   // ---------- 网络 7 ----------
   // 标题：Z06---> 摄像头防尘盖气缸
   // 注释：临时替换为RSP开关气缸
   // 含义：当 #ST01.Z06.RetEVT 为 TRUE 时置位 #ST01.Z06.IRetPos，否则复位（触点→线圈）
   IF #ST01.Z06.RetEVT THEN
       #ST01.Z06.IRetPos := TRUE;
   ELSE
       #ST01.Z06.IRetPos := FALSE;
   END_IF;
   // 含义：当 #ST01.Z06.ExtEVT 为 TRUE 时置位 #ST01.Z06.IExtPos，否则复位（触点→线圈）
   IF #ST01.Z06.ExtEVT THEN
       #ST01.Z06.IExtPos := TRUE;
   ELSE
       #ST01.Z06.IExtPos := FALSE;
   END_IF;
   // 含义：将 (NOT (#ST01.Z06.ExtEVT) AND #ST01.Z06.IRetPos) AND NOT (#ST01.Z06.IExtPos) 赋给 #ST01.Z06.RetPos
   #ST01.Z06.RetPos := (NOT (#ST01.Z06.ExtEVT) AND #ST01.Z06.IRetPos) AND NOT (#ST01.Z06.IExtPos);
   // 含义：将 (NOT (#ST01.Z06.ExtEVT) AND #ST01.Z06.IRetPos) AND NOT (#ST01.Z06.IExtPos) 赋给 "DB1900_Communication_PC".Send.Z06RetPos
   "DB1900_Communication_PC".Send.Z06RetPos := (NOT (#ST01.Z06.ExtEVT) AND #ST01.Z06.IRetPos) AND NOT (#ST01.Z06.IExtPos);
   // 含义：将 (NOT (#ST01.Z06.RetEVT) AND NOT (#ST01.Z06.IRetPos)) AND #ST01.Z06.IExtPos 赋给 #ST01.Z06.ExtPos
   #ST01.Z06.ExtPos := (NOT (#ST01.Z06.RetEVT) AND NOT (#ST01.Z06.IRetPos)) AND #ST01.Z06.IExtPos;
   // 含义：将 (NOT (#ST01.Z06.RetEVT) AND NOT (#ST01.Z06.IRetPos)) AND #ST01.Z06.IExtPos 赋给 "DB1900_Communication_PC".Send.Z06ExtPos
   "DB1900_Communication_PC".Send.Z06ExtPos := (NOT (#ST01.Z06.RetEVT) AND NOT (#ST01.Z06.IRetPos)) AND #ST01.Z06.IExtPos;
   // 含义：当 #OverAllPmt 为 TRUE 时置位 #ST01.Z06.ExtPmt，否则复位（触点→线圈）
   IF #OverAllPmt THEN
       #ST01.Z06.ExtPmt := TRUE;
   ELSE
       #ST01.Z06.ExtPmt := FALSE;
   END_IF;
   // 含义：当 #OverAllPmt 为 TRUE 时置位 #ST01.Z06.RetPmt，否则复位（触点→线圈）
   IF #OverAllPmt THEN
       #ST01.Z06.RetPmt := TRUE;
   ELSE
       #ST01.Z06.RetPmt := FALSE;
   END_IF;
   // 含义：调用块/实例 "DB1200_FB_std_Switch"，参数：CylinderCmd := #ST01.Z06
   "DB1200_FB_std_Switch"(CylinderCmd := #ST01.Z06);
   // 含义：当 #ST01.Z06.ExtIng 为 TRUE 时置位 "DB1146_PromptFree".ST01.Z06Exting，否则复位（触点→线圈）
   IF #ST01.Z06.ExtIng THEN
       "DB1146_PromptFree".ST01.Z06Exting := TRUE;
   ELSE
       "DB1146_PromptFree".ST01.Z06Exting := FALSE;
   END_IF;
   // 含义：当 #ST01.Z06.RetIng 为 TRUE 时置位 "DB1146_PromptFree".ST01.Z06Reting，否则复位（触点→线圈）
   IF #ST01.Z06.RetIng THEN
       "DB1146_PromptFree".ST01.Z06Reting := TRUE;
   ELSE
       "DB1146_PromptFree".ST01.Z06Reting := FALSE;
   END_IF;
   // 含义：当 #ST01.Z06.ExtErr 为 TRUE 时置位 "DB1148_PromptBeeper".ST01.Z06ExtErr，否则复位（触点→线圈）
   IF #ST01.Z06.ExtErr THEN
       "DB1148_PromptBeeper".ST01.Z06ExtErr := TRUE;
   ELSE
       "DB1148_PromptBeeper".ST01.Z06ExtErr := FALSE;
   END_IF;
   // 含义：当 #ST01.Z06.RetErr 为 TRUE 时置位 "DB1148_PromptBeeper".ST01.Z06RetErr，否则复位（触点→线圈）
   IF #ST01.Z06.RetErr THEN
       "DB1148_PromptBeeper".ST01.Z06RetErr := TRUE;
   ELSE
       "DB1148_PromptBeeper".ST01.Z06RetErr := FALSE;
   END_IF;
   // 含义：条件 "ManMode_M" AND "DB1900_Communication_PC".Recv.Z06ExtTPPB 成立时，将 TRUE 传送到 #ST01.Z06.ExtAuto
   IF "ManMode_M" AND "DB1900_Communication_PC".Recv.Z06ExtTPPB THEN
       #ST01.Z06.ExtAuto := TRUE;
   END_IF;
   // 含义：条件 "ManMode_M" AND "DB1900_Communication_PC".Recv.Z06RetTPPB 成立时，将 TRUE 传送到 #ST01.Z06.RetAuto
   IF "ManMode_M" AND "DB1900_Communication_PC".Recv.Z06RetTPPB THEN
       #ST01.Z06.RetAuto := TRUE;
   END_IF;

   // ---------- 网络 8 ----------
   // 标题：Z07--->快换盘锁紧
   // 含义：将 "IZ07RetPos" AND #Time.ST01Z07RET.Q 赋给 #ST01.Z07.IRetPos
   #ST01.Z07.IRetPos := "IZ07RetPos" AND #Time.ST01Z07RET.Q;
   // 含义：调用定时器实例 #Time.ST01Z07RET.TON
   #Time.ST01Z07RET.TON(IN := "IZ07RetPos",
                        PT := T#1S);
   // 含义：将 "IZ07ExtPos" AND #Time.ST01Z07EXT.Q 赋给 #ST01.Z07.IExtPos
   #ST01.Z07.IExtPos := "IZ07ExtPos" AND #Time.ST01Z07EXT.Q;
   // 含义：调用定时器实例 #Time.ST01Z07EXT.TON
   #Time.ST01Z07EXT.TON(IN := "IZ07ExtPos",
                        PT := T#1S);
   // 含义：将 (NOT (#ST01.Z07.ExtEVT) AND #ST01.Z07.IRetPos) AND NOT (#ST01.Z07.IExtPos) 赋给 #ST01.Z07.RetPos
   #ST01.Z07.RetPos := (NOT (#ST01.Z07.ExtEVT) AND #ST01.Z07.IRetPos) AND NOT (#ST01.Z07.IExtPos);
   // 含义：将 (NOT (#ST01.Z07.ExtEVT) AND #ST01.Z07.IRetPos) AND NOT (#ST01.Z07.IExtPos) 赋给 "DB1900_Communication_PC".Send.Z07RetPos
   "DB1900_Communication_PC".Send.Z07RetPos := (NOT (#ST01.Z07.ExtEVT) AND #ST01.Z07.IRetPos) AND NOT (#ST01.Z07.IExtPos);
   // 含义：将 (NOT (#ST01.Z07.RetEVT) AND NOT (#ST01.Z07.IRetPos)) AND #ST01.Z07.IExtPos 赋给 #ST01.Z07.ExtPos
   #ST01.Z07.ExtPos := (NOT (#ST01.Z07.RetEVT) AND NOT (#ST01.Z07.IRetPos)) AND #ST01.Z07.IExtPos;
   // 含义：将 (NOT (#ST01.Z07.RetEVT) AND NOT (#ST01.Z07.IRetPos)) AND #ST01.Z07.IExtPos 赋给 "DB1900_Communication_PC".Send.Z07ExtPos
   "DB1900_Communication_PC".Send.Z07ExtPos := (NOT (#ST01.Z07.RetEVT) AND NOT (#ST01.Z07.IRetPos)) AND #ST01.Z07.IExtPos;
   // 含义：将 (#OverAllPmt AND "DB720_KuKa_MainCtrl".StatusIn.do_ChgGrp_Pos) OR (#OverAllPmt AND TRUE) 赋给 #ST01.Z07.ExtPmt
   #ST01.Z07.ExtPmt := (#OverAllPmt AND "DB720_KuKa_MainCtrl".StatusIn.do_ChgGrp_Pos) OR (#OverAllPmt AND TRUE);
   // 含义：将 (#OverAllPmt AND "DB720_KuKa_MainCtrl".StatusIn.do_ChgGrp_Pos) OR (#OverAllPmt AND TRUE) 赋给 #ST01.Z07.RetPmt
   #ST01.Z07.RetPmt := (#OverAllPmt AND "DB720_KuKa_MainCtrl".StatusIn.do_ChgGrp_Pos) OR (#OverAllPmt AND TRUE);
   // 含义：调用块/实例 "DB1200_FB_std_Switch"，参数：CylinderCmd := #ST01.Z07
   "DB1200_FB_std_Switch"(CylinderCmd := #ST01.Z07);
   // 含义：当 #ST01.Z07.ExtIng 为 TRUE 时置位 "DB1146_PromptFree".ST01.Z07Exting，否则复位（触点→线圈）
   IF #ST01.Z07.ExtIng THEN
       "DB1146_PromptFree".ST01.Z07Exting := TRUE;
   ELSE
       "DB1146_PromptFree".ST01.Z07Exting := FALSE;
   END_IF;
   // 含义：当 #ST01.Z07.RetIng 为 TRUE 时置位 "DB1146_PromptFree".ST01.Z07Reting，否则复位（触点→线圈）
   IF #ST01.Z07.RetIng THEN
       "DB1146_PromptFree".ST01.Z07Reting := TRUE;
   ELSE
       "DB1146_PromptFree".ST01.Z07Reting := FALSE;
   END_IF;
   // 含义：当 #ST01.Z07.ExtErr 为 TRUE 时置位 "DB1148_PromptBeeper".ST01.Z07ExtErr，否则复位（触点→线圈）
   IF #ST01.Z07.ExtErr THEN
       "DB1148_PromptBeeper".ST01.Z07ExtErr := TRUE;
   ELSE
       "DB1148_PromptBeeper".ST01.Z07ExtErr := FALSE;
   END_IF;
   // 含义：当 #ST01.Z07.RetErr 为 TRUE 时置位 "DB1148_PromptBeeper".ST01.Z07RetErr，否则复位（触点→线圈）
   IF #ST01.Z07.RetErr THEN
       "DB1148_PromptBeeper".ST01.Z07RetErr := TRUE;
   ELSE
       "DB1148_PromptBeeper".ST01.Z07RetErr := FALSE;
   END_IF;
   // 含义：当 #ST01.Z07.ExtEVT 为 TRUE 时置位 "QZ07ExtEvt"，否则复位（触点→线圈）
   IF #ST01.Z07.ExtEVT THEN
       "QZ07ExtEvt" := TRUE;
   ELSE
       "QZ07ExtEvt" := FALSE;
   END_IF;
   // 含义：当 #ST01.Z07.RetEVT 为 TRUE 时置位 "QZ07RetEvt"，否则复位（触点→线圈）
   IF #ST01.Z07.RetEVT THEN
       "QZ07RetEvt" := TRUE;
   ELSE
       "QZ07RetEvt" := FALSE;
   END_IF;
   // 含义：条件 "ManMode_M" AND "DB1900_Communication_PC".Recv.Z07RetTPPB 成立时，将 TRUE 传送到 #ST01.Z07.RetAuto
   IF "ManMode_M" AND "DB1900_Communication_PC".Recv.Z07RetTPPB THEN
       #ST01.Z07.RetAuto := TRUE;
   END_IF;
   // 含义：条件 "ManMode_M" AND "DB1900_Communication_PC".Recv.Z07ExtTPPB 成立时，将 TRUE 传送到 #ST01.Z07.ExtAuto
   IF "ManMode_M" AND "DB1900_Communication_PC".Recv.Z07ExtTPPB THEN
       #ST01.Z07.ExtAuto := TRUE;
   END_IF;

   // ---------- 网络 9 ----------
   // 标题：Z08--->参数写入
   // 含义：将 #ST01.Z08.RetEVT AND #Time.ST01Z08RET.Q 赋给 #ST01.Z08.IRetPos
   #ST01.Z08.IRetPos := #ST01.Z08.RetEVT AND #Time.ST01Z08RET.Q;
   // 含义：调用定时器实例 #Time.ST01Z08RET.TON
   #Time.ST01Z08RET.TON(IN := #ST01.Z08.RetEVT,
                        PT := T#1S);
   // 含义：将 #ST01.Z08.ExtEVT AND #Time.ST01Z08EXT.Q 赋给 #ST01.Z08.IExtPos
   #ST01.Z08.IExtPos := #ST01.Z08.ExtEVT AND #Time.ST01Z08EXT.Q;
   // 含义：调用定时器实例 #Time.ST01Z08EXT.TON
   #Time.ST01Z08EXT.TON(IN := #ST01.Z08.ExtEVT,
                        PT := T#1S);
   // 含义：将 (NOT (#ST01.Z08.ExtEVT) AND #ST01.Z08.IRetPos) AND NOT (#ST01.Z08.IExtPos) 赋给 #ST01.Z08.RetPos
   #ST01.Z08.RetPos := (NOT (#ST01.Z08.ExtEVT) AND #ST01.Z08.IRetPos) AND NOT (#ST01.Z08.IExtPos);
   // 含义：将 (NOT (#ST01.Z08.RetEVT) AND NOT (#ST01.Z08.IRetPos)) AND #ST01.Z08.IExtPos 赋给 #ST01.Z08.ExtPos
   #ST01.Z08.ExtPos := (NOT (#ST01.Z08.RetEVT) AND NOT (#ST01.Z08.IRetPos)) AND #ST01.Z08.IExtPos;
   // 含义：当 #OverAllPmt 为 TRUE 时置位 #ST01.Z08.ExtPmt，否则复位（触点→线圈）
   IF #OverAllPmt THEN
       #ST01.Z08.ExtPmt := TRUE;
   ELSE
       #ST01.Z08.ExtPmt := FALSE;
   END_IF;
   // 含义：当 #OverAllPmt 为 TRUE 时置位 #ST01.Z08.RetPmt，否则复位（触点→线圈）
   IF #OverAllPmt THEN
       #ST01.Z08.RetPmt := TRUE;
   ELSE
       #ST01.Z08.RetPmt := FALSE;
   END_IF;
   // 含义：调用块/实例 "DB1200_FB_std_Switch"，参数：CylinderCmd := #ST01.Z08
   "DB1200_FB_std_Switch"(CylinderCmd := #ST01.Z08);
   // 含义：当 #ST01.Z08.ExtIng 为 TRUE 时置位 "DB1146_PromptFree".ST01.Z08Exting，否则复位（触点→线圈）
   IF #ST01.Z08.ExtIng THEN
       "DB1146_PromptFree".ST01.Z08Exting := TRUE;
   ELSE
       "DB1146_PromptFree".ST01.Z08Exting := FALSE;
   END_IF;
   // 含义：当 #ST01.Z08.RetIng 为 TRUE 时置位 "DB1146_PromptFree".ST01.Z08Reting，否则复位（触点→线圈）
   IF #ST01.Z08.RetIng THEN
       "DB1146_PromptFree".ST01.Z08Reting := TRUE;
   ELSE
       "DB1146_PromptFree".ST01.Z08Reting := FALSE;
   END_IF;
   // 含义：当 #ST01.Z08.ExtErr 为 TRUE 时置位 "DB1148_PromptBeeper".ST01.Z08ExtErr，否则复位（触点→线圈）
   IF #ST01.Z08.ExtErr THEN
       "DB1148_PromptBeeper".ST01.Z08ExtErr := TRUE;
   ELSE
       "DB1148_PromptBeeper".ST01.Z08ExtErr := FALSE;
   END_IF;
   // 含义：当 #ST01.Z08.RetErr 为 TRUE 时置位 "DB1148_PromptBeeper".ST01.Z08RetErr，否则复位（触点→线圈）
   IF #ST01.Z08.RetErr THEN
       "DB1148_PromptBeeper".ST01.Z08RetErr := TRUE;
   ELSE
       "DB1148_PromptBeeper".ST01.Z08RetErr := FALSE;
   END_IF;
   // 含义：当 #ST01.Z08.ExtEVT 为 TRUE 时置位 "DB1900_Communication_PC".Send.ParaWrite，否则复位（触点→线圈）
   IF #ST01.Z08.ExtEVT THEN
       "DB1900_Communication_PC".Send.ParaWrite := TRUE;
   ELSE
       "DB1900_Communication_PC".Send.ParaWrite := FALSE;
   END_IF;
   // 含义：条件 "DB1900_Communication_PC".Recv.ParaWriteDone AND NOT ("ASMMode_M") 成立时，将 TRUE 传送到 #ST01.Z08.RetAuto
   IF "DB1900_Communication_PC".Recv.ParaWriteDone AND NOT ("ASMMode_M") THEN
       #ST01.Z08.RetAuto := TRUE;
   END_IF;
   // 含义：条件 NOT (TRUE) AND NOT ("AllMode_M") 成立时，将 TRUE 传送到 #ST01.Z08.RetAuto
   IF NOT (TRUE) AND NOT ("AllMode_M") THEN
       #ST01.Z08.RetAuto := TRUE;
   END_IF;

   // ---------- 网络 10 ----------
   // 标题：Z09--->三爪卡盘夹爪气缸
   // 含义：条件 (((((NOT (TRUE) AND "AutoMode_M") AND "DB1900_Communication_PC".Para.DrillDirection1) OR ((NOT (TRUE) AND "AutoMode_M") AND "DB1900_Communication_PC".Para.DrillDirection3)) AND NOT ("DB1900_Communication_PC".Para.ProduceMode3)) OR (((((NOT (TRUE) AND "AutoMode_M") AND "DB1900_Communication_PC".Para.DrillDirection1) OR ((NOT (TRUE) AND "AutoMode_M") AND "DB1900_Communication_PC".Para.DrillDirection3)) AND "DB1900_Communication_PC".Para.ProduceMode3) AND "DB1060_AutoStep".HorDrillAutoStep.HorDrillStep.StopDrill_End) OR (((((NOT (TRUE) AND "AutoMode_M") AND "DB1900_Communication_PC".Para.DrillDirection1) OR ((NOT (TRUE) AND "AutoMode_M") AND "DB1900_Communication_PC".Para.DrillDirection3)) AND "DB1900_Communication_PC".Para.ProduceMode3) AND "DB1060_AutoStep".DownDrillAutoStep.DownDrillStep.StopDrill_End)) AND "DB720_KuKa_MainCtrl".Aux.ToolAtPosTimer.Q 成立时，将 TRUE 传送到 #ST01.Z09.ExtEVT
   IF (((((NOT (TRUE) AND "AutoMode_M") AND "DB1900_Communication_PC".Para.DrillDirection1) OR ((NOT (TRUE) AND "AutoMode_M") AND "DB1900_Communication_PC".Para.DrillDirection3)) AND NOT ("DB1900_Communication_PC".Para.ProduceMode3)) OR (((((NOT (TRUE) AND "AutoMode_M") AND "DB1900_Communication_PC".Para.DrillDirection1) OR ((NOT (TRUE) AND "AutoMode_M") AND "DB1900_Communication_PC".Para.DrillDirection3)) AND "DB1900_Communication_PC".Para.ProduceMode3) AND "DB1060_AutoStep".HorDrillAutoStep.HorDrillStep.StopDrill_End) OR (((((NOT (TRUE) AND "AutoMode_M") AND "DB1900_Communication_PC".Para.DrillDirection1) OR ((NOT (TRUE) AND "AutoMode_M") AND "DB1900_Communication_PC".Para.DrillDirection3)) AND "DB1900_Communication_PC".Para.ProduceMode3) AND "DB1060_AutoStep".DownDrillAutoStep.DownDrillStep.StopDrill_End)) AND "DB720_KuKa_MainCtrl".Aux.ToolAtPosTimer.Q THEN
       #ST01.Z09.ExtEVT := TRUE;
   END_IF;
   // 含义：条件 (((((NOT (TRUE) AND "AutoMode_M") AND "DB1900_Communication_PC".Para.DrillDirection1) OR ((NOT (TRUE) AND "AutoMode_M") AND "DB1900_Communication_PC".Para.DrillDirection3)) AND NOT ("DB1900_Communication_PC".Para.ProduceMode3)) OR (((((NOT (TRUE) AND "AutoMode_M") AND "DB1900_Communication_PC".Para.DrillDirection1) OR ((NOT (TRUE) AND "AutoMode_M") AND "DB1900_Communication_PC".Para.DrillDirection3)) AND "DB1900_Communication_PC".Para.ProduceMode3) AND "DB1060_AutoStep".HorDrillAutoStep.HorDrillStep.StopDrill_End) OR (((((NOT (TRUE) AND "AutoMode_M") AND "DB1900_Communication_PC".Para.DrillDirection1) OR ((NOT (TRUE) AND "AutoMode_M") AND "DB1900_Communication_PC".Para.DrillDirection3)) AND "DB1900_Communication_PC".Para.ProduceMode3) AND "DB1060_AutoStep".DownDrillAutoStep.DownDrillStep.StopDrill_End)) AND "DB720_KuKa_MainCtrl".Aux.ToolAtPosTimer.Q 成立时，将 FALSE 传送到 #ST01.Z09.RetEVT
   IF (((((NOT (TRUE) AND "AutoMode_M") AND "DB1900_Communication_PC".Para.DrillDirection1) OR ((NOT (TRUE) AND "AutoMode_M") AND "DB1900_Communication_PC".Para.DrillDirection3)) AND NOT ("DB1900_Communication_PC".Para.ProduceMode3)) OR (((((NOT (TRUE) AND "AutoMode_M") AND "DB1900_Communication_PC".Para.DrillDirection1) OR ((NOT (TRUE) AND "AutoMode_M") AND "DB1900_Communication_PC".Para.DrillDirection3)) AND "DB1900_Communication_PC".Para.ProduceMode3) AND "DB1060_AutoStep".HorDrillAutoStep.HorDrillStep.StopDrill_End) OR (((((NOT (TRUE) AND "AutoMode_M") AND "DB1900_Communication_PC".Para.DrillDirection1) OR ((NOT (TRUE) AND "AutoMode_M") AND "DB1900_Communication_PC".Para.DrillDirection3)) AND "DB1900_Communication_PC".Para.ProduceMode3) AND "DB1060_AutoStep".DownDrillAutoStep.DownDrillStep.StopDrill_End)) AND "DB720_KuKa_MainCtrl".Aux.ToolAtPosTimer.Q THEN
       #ST01.Z09.RetEVT := FALSE;
   END_IF;
   // 含义：调用计数器实例 #Time.ST01Z09EXT.TON（上升沿计数，当前值写入 CV）
   #Time.ST01Z09EXT.TON(IN := (((((((NOT (TRUE) AND "AutoMode_M") AND "DB1900_Communication_PC".Para.DrillDirection1) OR ((NOT (TRUE) AND "AutoMode_M") AND "DB1900_Communication_PC".Para.DrillDirection3)) AND "DB1900_Communication_PC".Para.ProduceMode3) AND "DB720_KuKa_MainCtrl".StatusIn.do_Gouge_Pos) OR (((((NOT (TRUE) AND "AutoMode_M") AND "DB1900_Communication_PC".Para.DrillDirection1) OR ((NOT (TRUE) AND "AutoMode_M") AND "DB1900_Communication_PC".Para.DrillDirection3)) AND "DB1900_Communication_PC".Para.ProduceMode3) AND "DB720_KuKa_MainCtrl".StatusIn.do_DownDril_Pos)) AND ("DB1900_Communication_PC".Recv.Current_2 >= "DB1900_Communication_PC".Para.CurrentMinLimit)),
                        PT := T#30ms);
   // 含义：条件 ((((((NOT (TRUE) AND "AutoMode_M") AND "DB1900_Communication_PC".Para.DrillDirection1) OR ((NOT (TRUE) AND "AutoMode_M") AND "DB1900_Communication_PC".Para.DrillDirection3)) AND "DB1900_Communication_PC".Para.ProduceMode3) AND "DB720_KuKa_MainCtrl".StatusIn.do_Gouge_Pos) OR (((((NOT (TRUE) AND "AutoMode_M") AND "DB1900_Communication_PC".Para.DrillDirection1) OR ((NOT (TRUE) AND "AutoMode_M") AND "DB1900_Communication_PC".Para.DrillDirection3)) AND "DB1900_Communication_PC".Para.ProduceMode3) AND "DB720_KuKa_MainCtrl".StatusIn.do_DownDril_Pos)) AND #Time.ST01Z09EXT.Q 成立时，将 FALSE 传送到 #ST01.Z09.ExtEVT
   IF ((((((NOT (TRUE) AND "AutoMode_M") AND "DB1900_Communication_PC".Para.DrillDirection1) OR ((NOT (TRUE) AND "AutoMode_M") AND "DB1900_Communication_PC".Para.DrillDirection3)) AND "DB1900_Communication_PC".Para.ProduceMode3) AND "DB720_KuKa_MainCtrl".StatusIn.do_Gouge_Pos) OR (((((NOT (TRUE) AND "AutoMode_M") AND "DB1900_Communication_PC".Para.DrillDirection1) OR ((NOT (TRUE) AND "AutoMode_M") AND "DB1900_Communication_PC".Para.DrillDirection3)) AND "DB1900_Communication_PC".Para.ProduceMode3) AND "DB720_KuKa_MainCtrl".StatusIn.do_DownDril_Pos)) AND #Time.ST01Z09EXT.Q THEN
       #ST01.Z09.ExtEVT := FALSE;
   END_IF;
   // 含义：条件 ((((((NOT (TRUE) AND "AutoMode_M") AND "DB1900_Communication_PC".Para.DrillDirection1) OR ((NOT (TRUE) AND "AutoMode_M") AND "DB1900_Communication_PC".Para.DrillDirection3)) AND "DB1900_Communication_PC".Para.ProduceMode3) AND "DB720_KuKa_MainCtrl".StatusIn.do_Gouge_Pos) OR (((((NOT (TRUE) AND "AutoMode_M") AND "DB1900_Communication_PC".Para.DrillDirection1) OR ((NOT (TRUE) AND "AutoMode_M") AND "DB1900_Communication_PC".Para.DrillDirection3)) AND "DB1900_Communication_PC".Para.ProduceMode3) AND "DB720_KuKa_MainCtrl".StatusIn.do_DownDril_Pos)) AND #Time.ST01Z09EXT.Q 成立时，将 TRUE 传送到 #ST01.Z09.RetEVT
   IF ((((((NOT (TRUE) AND "AutoMode_M") AND "DB1900_Communication_PC".Para.DrillDirection1) OR ((NOT (TRUE) AND "AutoMode_M") AND "DB1900_Communication_PC".Para.DrillDirection3)) AND "DB1900_Communication_PC".Para.ProduceMode3) AND "DB720_KuKa_MainCtrl".StatusIn.do_Gouge_Pos) OR (((((NOT (TRUE) AND "AutoMode_M") AND "DB1900_Communication_PC".Para.DrillDirection1) OR ((NOT (TRUE) AND "AutoMode_M") AND "DB1900_Communication_PC".Para.DrillDirection3)) AND "DB1900_Communication_PC".Para.ProduceMode3) AND "DB720_KuKa_MainCtrl".StatusIn.do_DownDril_Pos)) AND #Time.ST01Z09EXT.Q THEN
       #ST01.Z09.RetEVT := TRUE;
   END_IF;
   // 含义：条件 ((((NOT (TRUE) AND "AutoMode_M") AND "DB1900_Communication_PC".Para.DrillDirection1) OR ((NOT (TRUE) AND "AutoMode_M") AND "DB1900_Communication_PC".Para.DrillDirection3)) AND "DB1900_Communication_PC".Para.ProduceMode3) AND #ST01.Z09.ExtEVT 成立时，将 TRUE 传送到 "QZ14ExtEvt"
   IF ((((NOT (TRUE) AND "AutoMode_M") AND "DB1900_Communication_PC".Para.DrillDirection1) OR ((NOT (TRUE) AND "AutoMode_M") AND "DB1900_Communication_PC".Para.DrillDirection3)) AND "DB1900_Communication_PC".Para.ProduceMode3) AND #ST01.Z09.ExtEVT THEN
       "QZ14ExtEvt" := TRUE;
   END_IF;
   // 含义：条件 ((((NOT (TRUE) AND "AutoMode_M") AND "DB1900_Communication_PC".Para.DrillDirection1) OR ((NOT (TRUE) AND "AutoMode_M") AND "DB1900_Communication_PC".Para.DrillDirection3)) AND "DB1900_Communication_PC".Para.ProduceMode3) AND #ST01.Z09.ExtEVT 成立时，将 FALSE 传送到 "QZ14RetEvt"
   IF ((((NOT (TRUE) AND "AutoMode_M") AND "DB1900_Communication_PC".Para.DrillDirection1) OR ((NOT (TRUE) AND "AutoMode_M") AND "DB1900_Communication_PC".Para.DrillDirection3)) AND "DB1900_Communication_PC".Para.ProduceMode3) AND #ST01.Z09.ExtEVT THEN
       "QZ14RetEvt" := FALSE;
   END_IF;
   // 含义：条件 ((((NOT (TRUE) AND "AutoMode_M") AND "DB1900_Communication_PC".Para.DrillDirection1) OR ((NOT (TRUE) AND "AutoMode_M") AND "DB1900_Communication_PC".Para.DrillDirection3)) AND "DB1900_Communication_PC".Para.ProduceMode3) AND #ST01.Z09.RetEVT 成立时，将 FALSE 传送到 "QZ14ExtEvt"
   IF ((((NOT (TRUE) AND "AutoMode_M") AND "DB1900_Communication_PC".Para.DrillDirection1) OR ((NOT (TRUE) AND "AutoMode_M") AND "DB1900_Communication_PC".Para.DrillDirection3)) AND "DB1900_Communication_PC".Para.ProduceMode3) AND #ST01.Z09.RetEVT THEN
       "QZ14ExtEvt" := FALSE;
   END_IF;
   // 含义：条件 ((((NOT (TRUE) AND "AutoMode_M") AND "DB1900_Communication_PC".Para.DrillDirection1) OR ((NOT (TRUE) AND "AutoMode_M") AND "DB1900_Communication_PC".Para.DrillDirection3)) AND "DB1900_Communication_PC".Para.ProduceMode3) AND #ST01.Z09.RetEVT 成立时，将 TRUE 传送到 "QZ14RetEvt"
   IF ((((NOT (TRUE) AND "AutoMode_M") AND "DB1900_Communication_PC".Para.DrillDirection1) OR ((NOT (TRUE) AND "AutoMode_M") AND "DB1900_Communication_PC".Para.DrillDirection3)) AND "DB1900_Communication_PC".Para.ProduceMode3) AND #ST01.Z09.RetEVT THEN
       "QZ14RetEvt" := TRUE;
   END_IF;
   // 含义：条件 (NOT (TRUE) AND "ManMode_M") OR ((NOT (TRUE) AND "AutoMode_M") AND NOT ("DB1900_Communication_PC".Send.DrillRunning)) 成立时，将 FALSE 传送到 #ST01.Z09.ExtEVT
   IF (NOT (TRUE) AND "ManMode_M") OR ((NOT (TRUE) AND "AutoMode_M") AND NOT ("DB1900_Communication_PC".Send.DrillRunning)) THEN
       #ST01.Z09.ExtEVT := FALSE;
   END_IF;
   // 含义：条件 (NOT (TRUE) AND "ManMode_M") OR ((NOT (TRUE) AND "AutoMode_M") AND NOT ("DB1900_Communication_PC".Send.DrillRunning)) 成立时，将 FALSE 传送到 #ST01.Z09.RetEVT
   IF (NOT (TRUE) AND "ManMode_M") OR ((NOT (TRUE) AND "AutoMode_M") AND NOT ("DB1900_Communication_PC".Send.DrillRunning)) THEN
       #ST01.Z09.RetEVT := FALSE;
   END_IF;

   // ---------- 网络 11 ----------
   // （空白网络）
END_FUNCTION_BLOCK

FUNCTION_BLOCK "FB1910_DrillData"   // FB1910, SCL
{ S7_Optimized_Access := 'TRUE' }
// ============================================================
//  Block: FB1910_DrillData
//  ============================================================
//  编号：FB1910
//  原始语言：LAD（规则翻译为 SCL）
//  含义：Hammer
   VAR
      HorDrill : "UDT_DrillData";   // 水平水泥数据
      DownDrill : "UDT_DrillData";   // 垂直向下水泥数据
      AUX : Struct   // 静态变量
         LayerNo : Int := 1;   // 层数记忆
         HDirection : Int := 1;   // 水平方向1正2负
         DDirection : Int := 1;   // 向下方向1正2负
         GougeDrillWidth : Real;   // 凿击宽度要加10
      END_STRUCT;
      EdgeDetc : Struct   // 静态变量
         Pulse : Array[0..15] of Bool;   // 静态变量
      END_STRUCT;
      CurrentDrillWidth : Real;   // 静态变量
      CurrentDrillLength : Real;   // 静态变量
      CurrentDrillDepth : Real;   // 静态变量
      LastDrillWidth : Real;   // 静态变量
      LastDrillDepth : Real;   // 静态变量
      AlreadyDrillWidth : Real;   // 静态变量
      AlreadyDrillLength : Real;   // 静态变量
      MaxWidth : Real;   // 静态变量
      gi_OffsetX : Real;   // 静态变量
      gi_OffSetY : Real;   // 静态变量
      gi_OffSetZ : Real;   // 静态变量
      SlabWidth : Real := 0.0;   // 静态变量
      SlabLength : Real := 0.0;   // 静态变量
      PosNo : Int;   // 静态变量
      OppositeStartPos : Real;   // 静态变量
   END_VAR
   VAR_TEMP
      HorPosMod : Int;   // 临时变量
      DownPosMod : Int;   // 临时变量
   END_VAR
BEGIN

   // ---------- 网络 1 ----------
   // 标题：水泥长宽输入
   // 含义：条件 ((("DB1900_Communication_PC".Para.HorConcreteZ > 100.0) AND ("DB720_KuKa_MainCtrl".CmdOut.gi_ToolTypeNo = 2))) OR ((("DB1900_Communication_PC".Para.HorConcreteZ > 100.0) AND ("DB720_KuKa_MainCtrl".CmdOut.gi_ToolTypeNo = 18))) 成立时，将 "DB1900_Communication_PC".Para.HorConcreteZ 传送到 #HorDrill.SlabWidth
   IF ((("DB1900_Communication_PC".Para.HorConcreteZ > 100.0) AND ("DB720_KuKa_MainCtrl".CmdOut.gi_ToolTypeNo = 2))) OR ((("DB1900_Communication_PC".Para.HorConcreteZ > 100.0) AND ("DB720_KuKa_MainCtrl".CmdOut.gi_ToolTypeNo = 18))) THEN
       #HorDrill.SlabWidth := "DB1900_Communication_PC".Para.HorConcreteZ;
   END_IF;
   // 含义：条件 (((("DB1900_Communication_PC".Para.HorConcreteZ > 100.0) AND ("DB720_KuKa_MainCtrl".CmdOut.gi_ToolTypeNo = 13))) AND ("DB1900_Communication_PC".Para.Classification = 1)) 成立时，将 500.0 传送到 #HorDrill.SlabWidth
   IF (((("DB1900_Communication_PC".Para.HorConcreteZ > 100.0) AND ("DB720_KuKa_MainCtrl".CmdOut.gi_ToolTypeNo = 13))) AND ("DB1900_Communication_PC".Para.Classification = 1)) THEN
       #HorDrill.SlabWidth := 500.0;
   END_IF;
   // 含义：条件 ((((("DB1900_Communication_PC".Para.HorConcreteZ > 100.0) AND ("DB720_KuKa_MainCtrl".CmdOut.gi_ToolTypeNo = 13))) AND ("DB1900_Communication_PC".Para.Classification = 2))) OR ((((("DB1900_Communication_PC".Para.HorConcreteZ > 100.0) AND ("DB720_KuKa_MainCtrl".CmdOut.gi_ToolTypeNo = 13))) AND ("DB1900_Communication_PC".Para.Classification = 3))) 成立时，将 850.0 传送到 #HorDrill.SlabWidth
   IF ((((("DB1900_Communication_PC".Para.HorConcreteZ > 100.0) AND ("DB720_KuKa_MainCtrl".CmdOut.gi_ToolTypeNo = 13))) AND ("DB1900_Communication_PC".Para.Classification = 2))) OR ((((("DB1900_Communication_PC".Para.HorConcreteZ > 100.0) AND ("DB720_KuKa_MainCtrl".CmdOut.gi_ToolTypeNo = 13))) AND ("DB1900_Communication_PC".Para.Classification = 3))) THEN
       #HorDrill.SlabWidth := 850.0;
   END_IF;
   // 含义：条件 ((("DB1900_Communication_PC".Para.HorConcreteY > 200.0) AND ("DB720_KuKa_MainCtrl".CmdOut.gi_ToolTypeNo = 2))) OR ((("DB1900_Communication_PC".Para.HorConcreteY > 200.0) AND ("DB720_KuKa_MainCtrl".CmdOut.gi_ToolTypeNo = 18))) 成立时，将 "DB1900_Communication_PC".Para.HorConcreteY 传送到 #HorDrill.SlabLength
   IF ((("DB1900_Communication_PC".Para.HorConcreteY > 200.0) AND ("DB720_KuKa_MainCtrl".CmdOut.gi_ToolTypeNo = 2))) OR ((("DB1900_Communication_PC".Para.HorConcreteY > 200.0) AND ("DB720_KuKa_MainCtrl".CmdOut.gi_ToolTypeNo = 18))) THEN
       #HorDrill.SlabLength := "DB1900_Communication_PC".Para.HorConcreteY;
   END_IF;
   // 含义：条件 (((("DB1900_Communication_PC".Para.HorConcreteY > 200.0) AND ("DB720_KuKa_MainCtrl".CmdOut.gi_ToolTypeNo = 13))) AND ("DB1900_Communication_PC".Para.DrillWidth <> 105.0)) 成立时，将 960.0 传送到 #HorDrill.SlabLength
   IF (((("DB1900_Communication_PC".Para.HorConcreteY > 200.0) AND ("DB720_KuKa_MainCtrl".CmdOut.gi_ToolTypeNo = 13))) AND ("DB1900_Communication_PC".Para.DrillWidth <> 105.0)) THEN
       #HorDrill.SlabLength := 960.0;
   END_IF;
   // 含义：条件 (((("DB1900_Communication_PC".Para.HorConcreteY > 200.0) AND ("DB720_KuKa_MainCtrl".CmdOut.gi_ToolTypeNo = 13))) AND ("DB1900_Communication_PC".Para.DrillWidth = 105.0)) 成立时，将 1100.0 传送到 #HorDrill.SlabLength
   IF (((("DB1900_Communication_PC".Para.HorConcreteY > 200.0) AND ("DB720_KuKa_MainCtrl".CmdOut.gi_ToolTypeNo = 13))) AND ("DB1900_Communication_PC".Para.DrillWidth = 105.0)) THEN
       #HorDrill.SlabLength := 1100.0;
   END_IF;
   // 含义：条件 ("DB1900_Communication_PC".Para.DownConcreteX > 50.0) 成立时，将 "DB1900_Communication_PC".Para.DownConcreteX 传送到 #DownDrill.SlabWidth
   IF ("DB1900_Communication_PC".Para.DownConcreteX > 50.0) THEN
       #DownDrill.SlabWidth := "DB1900_Communication_PC".Para.DownConcreteX;
   END_IF;
   // 含义：条件 (("DB1900_Communication_PC".Para.DownConcreteY > 100.0) AND ("DB720_KuKa_MainCtrl".CmdOut.gi_ToolTypeNo = 2)) 成立时，将 "DB1900_Communication_PC".Para.DownConcreteY 传送到 #DownDrill.SlabLength
   IF (("DB1900_Communication_PC".Para.DownConcreteY > 100.0) AND ("DB720_KuKa_MainCtrl".CmdOut.gi_ToolTypeNo = 2)) THEN
       #DownDrill.SlabLength := "DB1900_Communication_PC".Para.DownConcreteY;
   END_IF;
   // 含义：条件 (("DB1900_Communication_PC".Para.DownConcreteY > 100.0) AND ("DB720_KuKa_MainCtrl".CmdOut.gi_ToolTypeNo = 13)) 成立时，将 1110.0 传送到 #DownDrill.SlabLength
   IF (("DB1900_Communication_PC".Para.DownConcreteY > 100.0) AND ("DB720_KuKa_MainCtrl".CmdOut.gi_ToolTypeNo = 13)) THEN
       #DownDrill.SlabLength := 1110.0;
   END_IF;
   // 含义：条件 ("DB1900_Communication_PC".Recv.Layer < 1) 成立时，将 1 传送到 "DB1900_Communication_PC".Recv.Layer
   IF ("DB1900_Communication_PC".Recv.Layer < 1) THEN
       "DB1900_Communication_PC".Recv.Layer := 1;
   END_IF;
   // 含义：条件 "DB1900_Communication_PC".Recv.PowerOff OR ("ManMode_M" AND "ErrRst_M") 成立时，将 FALSE 传送到 "DB1900_Communication_PC".Send.PowerOff
   IF "DB1900_Communication_PC".Recv.PowerOff OR ("ManMode_M" AND "ErrRst_M") THEN
       "DB1900_Communication_PC".Send.PowerOff := FALSE;
   END_IF;

   // ---------- 网络 2 ----------
   // 标题：锤钻打孔长宽输入
   // 注释：Hammer
   // 含义：条件 ((("DB720_KuKa_MainCtrl".CmdOut.gi_ToolTypeNo = 2) OR ("DB720_KuKa_MainCtrl".CmdOut.gi_ToolTypeNo = 18)) AND "DB1900_Communication_PC".Para.DrillDirection1) AND NOT ("DB1900_Communication_PC".Para.ProduceMode3) 成立时，将 "DB1900_Communication_PC".Para.DrillWidth 传送到 #HorDrill.CurrentDrillWidth
   IF ((("DB720_KuKa_MainCtrl".CmdOut.gi_ToolTypeNo = 2) OR ("DB720_KuKa_MainCtrl".CmdOut.gi_ToolTypeNo = 18)) AND "DB1900_Communication_PC".Para.DrillDirection1) AND NOT ("DB1900_Communication_PC".Para.ProduceMode3) THEN
       #HorDrill.CurrentDrillWidth := "DB1900_Communication_PC".Para.DrillWidth;
   END_IF;
   // 含义：条件 ((("DB720_KuKa_MainCtrl".CmdOut.gi_ToolTypeNo = 2) OR ("DB720_KuKa_MainCtrl".CmdOut.gi_ToolTypeNo = 18)) AND "DB1900_Communication_PC".Para.DrillDirection1) AND "DB1900_Communication_PC".Para.ProduceMode3 成立时，将 ("DB1900_Communication_PC".Para.DrillWidth + 10.0) 传送到 #HorDrill.CurrentDrillWidth
   IF ((("DB720_KuKa_MainCtrl".CmdOut.gi_ToolTypeNo = 2) OR ("DB720_KuKa_MainCtrl".CmdOut.gi_ToolTypeNo = 18)) AND "DB1900_Communication_PC".Para.DrillDirection1) AND "DB1900_Communication_PC".Para.ProduceMode3 THEN
       #HorDrill.CurrentDrillWidth := ("DB1900_Communication_PC".Para.DrillWidth + 10.0);
   END_IF;
   // 含义：条件 (("DB720_KuKa_MainCtrl".CmdOut.gi_ToolTypeNo = 2) OR ("DB720_KuKa_MainCtrl".CmdOut.gi_ToolTypeNo = 18)) AND "DB1900_Communication_PC".Para.DrillDirection1 成立时，将 "DB1900_Communication_PC".Para.DrillWidth 传送到 #HorDrill.CurrentDrillLength
   IF (("DB720_KuKa_MainCtrl".CmdOut.gi_ToolTypeNo = 2) OR ("DB720_KuKa_MainCtrl".CmdOut.gi_ToolTypeNo = 18)) AND "DB1900_Communication_PC".Para.DrillDirection1 THEN
       #HorDrill.CurrentDrillLength := "DB1900_Communication_PC".Para.DrillWidth;
   END_IF;
   // 含义：条件 (("DB720_KuKa_MainCtrl".CmdOut.gi_ToolTypeNo = 2) OR ("DB720_KuKa_MainCtrl".CmdOut.gi_ToolTypeNo = 18)) AND "DB1900_Communication_PC".Para.DrillDirection3 成立时，将 "DB1900_Communication_PC".Para.DrillWidth 传送到 #DownDrill.CurrentDrillWidth
   IF (("DB720_KuKa_MainCtrl".CmdOut.gi_ToolTypeNo = 2) OR ("DB720_KuKa_MainCtrl".CmdOut.gi_ToolTypeNo = 18)) AND "DB1900_Communication_PC".Para.DrillDirection3 THEN
       #DownDrill.CurrentDrillWidth := "DB1900_Communication_PC".Para.DrillWidth;
   END_IF;

   // ---------- 网络 3 ----------
   // 标题：打孔水钻长宽输入
   // 注释：Core Diamond Drill
   // 32mm: Hor; Height:  45mm; Length: 50mm 100mm   150mm 250mm
   // 52mm:Down; Height: 65mm; Length: 66.66mm 132.33mmmm   233.67mm
   // 82mm Hor; Height:85mm; Length:100mm 300mm
   // 102mm Hor; Height:80mm; Length:400mm
   // 132mm Hor; Height:120mm; Length:400mm
   // 含义：条件 ((((("DB720_KuKa_MainCtrl".CmdOut.gi_ToolTypeNo = 13) AND "DB1900_Communication_PC".Para.DrillDirection1) AND ("DB1900_Communication_PC".Para.DrillWidth = 45.0))) AND ("DB1900_Communication_PC".Para.Classification = 1)) 成立时，将 (#HorDrill.PosNo MOD 4) 传送到 #HorPosMod
   IF ((((("DB720_KuKa_MainCtrl".CmdOut.gi_ToolTypeNo = 13) AND "DB1900_Communication_PC".Para.DrillDirection1) AND ("DB1900_Communication_PC".Para.DrillWidth = 45.0))) AND ("DB1900_Communication_PC".Para.Classification = 1)) THEN
       #HorPosMod := (#HorDrill.PosNo MOD 4);
   END_IF;
   // 含义：条件 ((#HorDrill.PosNo >= 1) AND (#HorPosMod = 3)) 成立时，将 250.0 传送到 #HorDrill.CurrentDrillLength
   IF ((#HorDrill.PosNo >= 1) AND (#HorPosMod = 3)) THEN
       #HorDrill.CurrentDrillLength := 250.0;
   END_IF;
   // 含义：条件 ((#HorDrill.PosNo >= 1) AND (#HorPosMod <> 3)) 成立时，将 50.0 传送到 #HorDrill.CurrentDrillLength
   IF ((#HorDrill.PosNo >= 1) AND (#HorPosMod <> 3)) THEN
       #HorDrill.CurrentDrillLength := 50.0;
   END_IF;
   // 含义：条件 ((#HorDrill.PosNo = 0) AND (#HorPosMod = 0)) 成立时，将 50.0 传送到 #HorDrill.CurrentDrillLength
   IF ((#HorDrill.PosNo = 0) AND (#HorPosMod = 0)) THEN
       #HorDrill.CurrentDrillLength := 50.0;
   END_IF;
   // 含义：条件 ((((("DB720_KuKa_MainCtrl".CmdOut.gi_ToolTypeNo = 13) AND "DB1900_Communication_PC".Para.DrillDirection1) AND ("DB1900_Communication_PC".Para.DrillWidth = 65.0))) AND ("DB1900_Communication_PC".Para.Classification = 1)) 成立时，将 (#HorDrill.PosNo MOD 3) 传送到 #HorPosMod
   IF ((((("DB720_KuKa_MainCtrl".CmdOut.gi_ToolTypeNo = 13) AND "DB1900_Communication_PC".Para.DrillDirection1) AND ("DB1900_Communication_PC".Para.DrillWidth = 65.0))) AND ("DB1900_Communication_PC".Para.Classification = 1)) THEN
       #HorPosMod := (#HorDrill.PosNo MOD 3);
   END_IF;
   // 含义：条件 ((#HorDrill.PosNo >= 1) AND (#HorPosMod = 2)) 成立时，将 266.68 传送到 #HorDrill.CurrentDrillLength
   IF ((#HorDrill.PosNo >= 1) AND (#HorPosMod = 2)) THEN
       #HorDrill.CurrentDrillLength := 266.68;
   END_IF;
   // 含义：条件 ((#HorDrill.PosNo >= 1) AND (#HorPosMod <> 2)) 成立时，将 66.66 传送到 #HorDrill.CurrentDrillLength
   IF ((#HorDrill.PosNo >= 1) AND (#HorPosMod <> 2)) THEN
       #HorDrill.CurrentDrillLength := 66.66;
   END_IF;
   // 含义：条件 ((#HorDrill.PosNo = 0) AND (#HorPosMod = 0)) 成立时，将 66.66 传送到 #HorDrill.CurrentDrillLength
   IF ((#HorDrill.PosNo = 0) AND (#HorPosMod = 0)) THEN
       #HorDrill.CurrentDrillLength := 66.66;
   END_IF;
   // 含义：条件 (((((("DB720_KuKa_MainCtrl".CmdOut.gi_ToolTypeNo = 13) AND "DB1900_Communication_PC".Para.DrillDirection1) AND ("DB1900_Communication_PC".Para.DrillWidth = 85.0))) AND ("DB1900_Communication_PC".Para.Classification = 2))) OR (((((("DB720_KuKa_MainCtrl".CmdOut.gi_ToolTypeNo = 13) AND "DB1900_Communication_PC".Para.DrillDirection1) AND ("DB1900_Communication_PC".Para.DrillWidth = 85.0))) AND ("DB1900_Communication_PC".Para.Classification = 3))) 成立时，将 (#HorDrill.PosNo MOD 2) 传送到 #HorPosMod
   IF (((((("DB720_KuKa_MainCtrl".CmdOut.gi_ToolTypeNo = 13) AND "DB1900_Communication_PC".Para.DrillDirection1) AND ("DB1900_Communication_PC".Para.DrillWidth = 85.0))) AND ("DB1900_Communication_PC".Para.Classification = 2))) OR (((((("DB720_KuKa_MainCtrl".CmdOut.gi_ToolTypeNo = 13) AND "DB1900_Communication_PC".Para.DrillDirection1) AND ("DB1900_Communication_PC".Para.DrillWidth = 85.0))) AND ("DB1900_Communication_PC".Para.Classification = 3))) THEN
       #HorPosMod := (#HorDrill.PosNo MOD 2);
   END_IF;
   // 含义：条件 ((#HorDrill.PosNo >= 1) AND (#HorPosMod = 1)) 成立时，将 300.0 传送到 #HorDrill.CurrentDrillLength
   IF ((#HorDrill.PosNo >= 1) AND (#HorPosMod = 1)) THEN
       #HorDrill.CurrentDrillLength := 300.0;
   END_IF;
   // 含义：条件 ((#HorDrill.PosNo >= 1) AND (#HorPosMod <> 1)) 成立时，将 100.0 传送到 #HorDrill.CurrentDrillLength
   IF ((#HorDrill.PosNo >= 1) AND (#HorPosMod <> 1)) THEN
       #HorDrill.CurrentDrillLength := 100.0;
   END_IF;
   // 含义：条件 ((#HorDrill.PosNo = 0) AND (#HorPosMod = 0)) 成立时，将 100.0 传送到 #HorDrill.CurrentDrillLength
   IF ((#HorDrill.PosNo = 0) AND (#HorPosMod = 0)) THEN
       #HorDrill.CurrentDrillLength := 100.0;
   END_IF;
   // 含义：条件 ((((("DB720_KuKa_MainCtrl".CmdOut.gi_ToolTypeNo = 13) AND "DB1900_Communication_PC".Para.DrillDirection1) AND ("DB1900_Communication_PC".Para.DrillWidth = 105.0))) AND ("DB1900_Communication_PC".Para.Classification = 1)) 成立时，将 125.0 传送到 #HorDrill.CurrentDrillLength
   IF ((((("DB720_KuKa_MainCtrl".CmdOut.gi_ToolTypeNo = 13) AND "DB1900_Communication_PC".Para.DrillDirection1) AND ("DB1900_Communication_PC".Para.DrillWidth = 105.0))) AND ("DB1900_Communication_PC".Para.Classification = 1)) THEN
       #HorDrill.CurrentDrillLength := 125.0;
   END_IF;
   // 含义：条件 (((((("DB720_KuKa_MainCtrl".CmdOut.gi_ToolTypeNo = 13) AND "DB1900_Communication_PC".Para.DrillDirection1) AND ("DB1900_Communication_PC".Para.DrillWidth = 80.0))) OR (((("DB720_KuKa_MainCtrl".CmdOut.gi_ToolTypeNo = 13) AND "DB1900_Communication_PC".Para.DrillDirection1) AND ("DB1900_Communication_PC".Para.DrillWidth = 120.0)))) AND ("DB1900_Communication_PC".Para.Classification = 2)) 成立时，将 400.0 传送到 #HorDrill.CurrentDrillLength
   IF (((((("DB720_KuKa_MainCtrl".CmdOut.gi_ToolTypeNo = 13) AND "DB1900_Communication_PC".Para.DrillDirection1) AND ("DB1900_Communication_PC".Para.DrillWidth = 80.0))) OR (((("DB720_KuKa_MainCtrl".CmdOut.gi_ToolTypeNo = 13) AND "DB1900_Communication_PC".Para.DrillDirection1) AND ("DB1900_Communication_PC".Para.DrillWidth = 120.0)))) AND ("DB1900_Communication_PC".Para.Classification = 2)) THEN
       #HorDrill.CurrentDrillLength := 400.0;
   END_IF;
   // 含义：条件 ("DB720_KuKa_MainCtrl".CmdOut.gi_ToolTypeNo = 13) AND "DB1900_Communication_PC".Para.DrillDirection1 成立时，将 "DB1900_Communication_PC".Para.DrillWidth 传送到 #HorDrill.CurrentDrillWidth
   IF ("DB720_KuKa_MainCtrl".CmdOut.gi_ToolTypeNo = 13) AND "DB1900_Communication_PC".Para.DrillDirection1 THEN
       #HorDrill.CurrentDrillWidth := "DB1900_Communication_PC".Para.DrillWidth;
   END_IF;
   // 含义：条件 ((("DB720_KuKa_MainCtrl".CmdOut.gi_ToolTypeNo = 13) AND "DB1900_Communication_PC".Para.DrillDirection3) AND ("DB1900_Communication_PC".Para.DrillWidth = 65.0)) 成立时，将 (#DownDrill.PosNo MOD 3) 传送到 #DownPosMod
   IF ((("DB720_KuKa_MainCtrl".CmdOut.gi_ToolTypeNo = 13) AND "DB1900_Communication_PC".Para.DrillDirection3) AND ("DB1900_Communication_PC".Para.DrillWidth = 65.0)) THEN
       #DownPosMod := (#DownDrill.PosNo MOD 3);
   END_IF;
   // 含义：条件 ((#DownDrill.PosNo >= 1) AND (#DownPosMod = 2)) 成立时，将 266.68 传送到 #DownDrill.CurrentDrillLength
   IF ((#DownDrill.PosNo >= 1) AND (#DownPosMod = 2)) THEN
       #DownDrill.CurrentDrillLength := 266.68;
   END_IF;
   // 含义：条件 ((#DownDrill.PosNo >= 1) AND (#DownPosMod <> 2)) 成立时，将 66.6 传送到 #DownDrill.CurrentDrillLength
   IF ((#DownDrill.PosNo >= 1) AND (#DownPosMod <> 2)) THEN
       #DownDrill.CurrentDrillLength := 66.6;
   END_IF;
   // 含义：条件 ((#DownDrill.PosNo = 0) AND (#DownPosMod = 0)) 成立时，将 66.6 传送到 #HorDrill.CurrentDrillLength
   IF ((#DownDrill.PosNo = 0) AND (#DownPosMod = 0)) THEN
       #HorDrill.CurrentDrillLength := 66.6;
   END_IF;
   // 含义：条件 ("DB720_KuKa_MainCtrl".CmdOut.gi_ToolTypeNo = 13) AND "DB1900_Communication_PC".Para.DrillDirection3 成立时，将 "DB1900_Communication_PC".Para.DrillWidth 传送到 #DownDrill.CurrentDrillWidth
   IF ("DB720_KuKa_MainCtrl".CmdOut.gi_ToolTypeNo = 13) AND "DB1900_Communication_PC".Para.DrillDirection3 THEN
       #DownDrill.CurrentDrillWidth := "DB1900_Communication_PC".Para.DrillWidth;
   END_IF;

   // ---------- 网络 4 ----------
   // 标题：手动输入水平水泥数据处理
   // 含义：本网络为 StructuredText（SCL）原文重建，非 LAD 折叠
   IF "DB1900_Communication_PC".Recv.HorizontalConfirm AND "IMan" THEN
       #AUX.HDirection := 1;
       #HorDrill.OppositeStartPos := 0;
       #AUX.LayerNo := "DB1900_Communication_PC".Recv.Layer;
       #HorDrill.LastDrillWidth := #HorDrill.CurrentDrillWidth;
       #HorDrill.gi_OffSetZ := ABS("DB1900_Communication_PC".Recv.Horizontal_OffSetZ);
       #HorDrill.gi_OffSetY := ABS("DB1900_Communication_PC".Recv.Horizontal_OffSetY);
       #HorDrill.AlreadyDrillWidth := ABS("DB1900_Communication_PC".Recv.Horizontal_OffSetZ);
       #HorDrill.AlreadyDrillLength := ABS("DB1900_Communication_PC".Recv.Horizontal_OffSetY);
       IF "DB1900_Communication_PC".Recv.Horizontal_OffSetY = 0 THEN
           #HorDrill.PosNo := 0;
       END_IF;
   END_IF;
   IF "DB1900_Communication_PC".Recv.ChangeHorizontalSlabDone AND "IMan" THEN
       #AUX.LayerNo := 1;
       #AUX.HDirection := 1;
       #HorDrill.PosNo := 0;
       #HorDrill.gi_OffSetZ := 0;
       #HorDrill.gi_OffSetY := 0;
       #HorDrill.OppositeStartPos := 0;
       #HorDrill.AlreadyDrillWidth := 0;
       #HorDrill.AlreadyDrillLength := 0;
       #HorDrill.LastDrillWidth := #HorDrill.CurrentDrillWidth;
       "DB1147_PromptStartNotPmt".Public.ChangeHorDrillSlab := FALSE;
   END_IF;

   // ---------- 网络 5 ----------
   // 标题：水平水泥数据 Y平长 Z纵宽
   // 含义：本网络为 StructuredText（SCL）原文重建，非 LAD 折叠
   IF "DB1900_Communication_PC".Para.DrillDirection1 = TRUE AND (NOT "DB1900_Communication_PC".Para.ProduceMode3) AND "AutoMode_M" THEN
       IF "DB2500 Visual Chiseling".VChiselCamRound = -1 THEN
           #HorDrill.SlabWidth := #HorDrill.SlabWidth;
       ELSIF ("DB2500 Visual Chiseling".VChiselCamRound >= 0 AND "DB2500 Visual Chiseling".VChiselCamRound <= 44) OR
           ("DB2500 Visual Chiseling".CalCamRound_Mid >= 0 AND "DB2500 Visual Chiseling".CalCamRound_Mid <= 2) THEN
           #HorDrill.SlabWidth := #HorDrill.SlabWidth - 300 - 30;
       ELSIF ("DB2500 Visual Chiseling".VChiselCamRound >= 45 OR "DB2500 Visual Chiseling".CalCamRound_Mid >= 3) THEN
           #HorDrill.SlabWidth := #HorDrill.SlabWidth - 500 - 30;
       END_IF;
       IF (("DB720_KuKa_MainCtrl".CmdOut.gi_ToolTypeNo = 13 OR "DB720_KuKa_MainCtrl".CmdOut.gi_ToolTypeNo = 18) AND
           NOT "DB1060_AutoStep".HorDrillAutoStep.HorDrillStep.StepStart) OR
           "DB720_KuKa_MainCtrl".CmdOut.gi_ToolTypeNo = 2 THEN
           IF #HorDrill.gi_OffSetZ <= #HorDrill.SlabWidth THEN
               "DB1147_PromptStartNotPmt".Public.ChangeHorDrillSlab := FALSE;
               IF #HorDrill.AlreadyDrillLength > #HorDrill.SlabLength OR
                   ((#HorDrill.OppositeStartPos - #HorDrill.AlreadyDrillLength < 0) AND
                   #HorDrill.OppositeStartPos <> 0 AND #AUX.HDirection = 2)
               THEN
                   IF #HorDrill.AlreadyDrillLength <> 0 THEN
                       IF #HorDrill.AlreadyDrillLength > #HorDrill.SlabLength THEN
                           #HorDrill.OppositeStartPos := #HorDrill.SlabLength;
                       ELSE
                           #HorDrill.OppositeStartPos := #HorDrill.AlreadyDrillLength;
                       END_IF;
                   END_IF;
                   #HorDrill.PosNo := 0;
                   #HorDrill.AlreadyDrillLength := 0;
                   #HorDrill.gi_OffSetZ := (#HorDrill.AlreadyDrillWidth + #HorDrill.CurrentDrillWidth);
                   #HorDrill.AlreadyDrillWidth := (#HorDrill.CurrentDrillWidth + #HorDrill.AlreadyDrillWidth);
                   IF #AUX.HDirection = 1 THEN
                       #AUX.HDirection := 2;
                       IF "DB720_KuKa_MainCtrl".CmdOut.gi_ToolTypeNo = 2 OR "DB720_KuKa_MainCtrl".CmdOut.gi_ToolTypeNo = 18 THEN
                           IF #HorDrill.OppositeStartPos + #HorDrill.CurrentDrillLength / 2 > #HorDrill.SlabLength THEN
                               #HorDrill.OppositeStartPos := #HorDrill.OppositeStartPos - #HorDrill.CurrentDrillLength / 2;
                           ELSE
                               #HorDrill.OppositeStartPos := #HorDrill.OppositeStartPos + #HorDrill.CurrentDrillLength / 2;
                           END_IF;
                       END_IF;
                       IF "DB720_KuKa_MainCtrl".CmdOut.gi_ToolTypeNo = 13 THEN
                           IF "DB1900_Communication_PC".Para.DrillWidth = 120.0 OR
                               "DB1900_Communication_PC".Para.DrillWidth = 80.0 OR
                               "DB1900_Communication_PC".Para.DrillWidth = 65.0 THEN
                               #HorDrill.OppositeStartPos := 900.0;
                           ELSIF "DB1900_Communication_PC".Para.DrillWidth = 45 THEN
                               #HorDrill.OppositeStartPos := 925.0;
                           ELSIF "DB1900_Communication_PC".Para.DrillWidth = 85.0 THEN
                               #HorDrill.OppositeStartPos := 850.0;
                           ELSIF "DB1900_Communication_PC".Para.DrillWidth = 105.0 THEN
                               #HorDrill.OppositeStartPos := 1062.5;
                           END_IF;
                       END_IF;
                   ELSE
                       #AUX.HDirection := 1;
                       #HorDrill.gi_OffSetY := 0;
                       #HorDrill.OppositeStartPos := 0;
                   END_IF;
               ELSE
                   IF #AUX.HDirection = 1 THEN
                       #HorDrill.gi_OffSetY := #HorDrill.AlreadyDrillLength;
                   ELSE
                       #HorDrill.gi_OffSetY := #HorDrill.OppositeStartPos - #HorDrill.AlreadyDrillLength;
                   END_IF;
                   IF #HorDrill.CurrentDrillWidth <> #HorDrill.LastDrillWidth AND #HorDrill.PosNo <> 1 THEN
                       IF "DB720_KuKa_MainCtrl".CmdOut.gi_ToolTypeNo = 2 OR "DB720_KuKa_MainCtrl".CmdOut.gi_ToolTypeNo = 18 THEN
                           #HorDrill.AlreadyDrillWidth := #HorDrill.AlreadyDrillWidth + ABS(#HorDrill.CurrentDrillWidth / 2 - #HorDrill.LastDrillWidth / 2);
                       ELSIF "DB720_KuKa_MainCtrl".CmdOut.gi_ToolTypeNo = 13 THEN
                           #HorDrill.AlreadyDrillWidth := #HorDrill.AlreadyDrillWidth + ABS(#HorDrill.CurrentDrillWidth / 2 - #HorDrill.LastDrillWidth / 2) + 20;
                       END_IF;
                       #HorDrill.gi_OffSetZ := #HorDrill.AlreadyDrillWidth;
                       #HorDrill.LastDrillWidth := #HorDrill.CurrentDrillWidth;
                   END_IF;
               END_IF;
           ELSE
               "DB1900_Communication_PC".Send.PowerOff := TRUE;
               "DB1147_PromptStartNotPmt".Public.ChangeHorDrillSlab := TRUE;
           END_IF;
       END_IF;
   END_IF;

   // ---------- 网络 6 ----------
   // 标题：手动输入向下水泥数据处理
   // 含义：本网络为 StructuredText（SCL）原文重建，非 LAD 折叠
   IF "DB1900_Communication_PC".Recv.DownloadConfirm AND "IMan" THEN
       #AUX.DDirection := 1;
       #DownDrill.OppositeStartPos := 0;
       #AUX.LayerNo := "DB1900_Communication_PC".Recv.Layer;
       #DownDrill.LastDrillWidth := #DownDrill.CurrentDrillWidth;
       #DownDrill.gi_OffsetX := ABS("DB1900_Communication_PC".Recv.Download_OffSetX);
       #DownDrill.gi_OffSetY := ABS("DB1900_Communication_PC".Recv.Download_OffSetY);
       #DownDrill.AlreadyDrillWidth := ABS("DB1900_Communication_PC".Recv.Download_OffSetX);
       #DownDrill.AlreadyDrillLength := ABS("DB1900_Communication_PC".Recv.Download_OffSetY);
       IF "DB1900_Communication_PC".Recv.Download_OffSetY = 0 THEN
           #DownDrill.PosNo := 0;
       END_IF;
   END_IF;
   IF "DB1900_Communication_PC".Recv.ChangeDownloadSlabDone AND "IMan" THEN
       #AUX.DDirection := 1;
       #DownDrill.PosNo := 0;
       #DownDrill.gi_OffsetX := 0;
       #DownDrill.gi_OffSetY := 0;
       #DownDrill.OppositeStartPos := 0;
       #DownDrill.AlreadyDrillWidth := 0;
       #DownDrill.AlreadyDrillLength := 0;
       #DownDrill.LastDrillWidth := #DownDrill.CurrentDrillWidth;
       "DB1147_PromptStartNotPmt".Public.ChangeDownloadSlab := FALSE;
   END_IF;

   // ---------- 网络 7 ----------
   // 标题：向下水泥数据 Y平长 X纵宽
   // 含义：本网络为 StructuredText（SCL）原文重建，非 LAD 折叠
   IF "DB1900_Communication_PC".Para.DrillDirection3 = TRUE AND "AutoMode_M" THEN
       IF ("DB720_KuKa_MainCtrl".CmdOut.gi_ToolTypeNo = 13 AND NOT "DB1060_AutoStep".DownDrillAutoStep.DownDrillStep.StepStart) OR
           "DB720_KuKa_MainCtrl".CmdOut.gi_ToolTypeNo = 2 THEN
           IF #DownDrill.gi_OffsetX <= #DownDrill.SlabWidth THEN
               "DB1147_PromptStartNotPmt".Public.ChangeDownloadSlab := FALSE;
               IF #DownDrill.AlreadyDrillLength > #DownDrill.SlabLength OR
                   ((#DownDrill.OppositeStartPos - #DownDrill.AlreadyDrillLength < 0) AND
                   #DownDrill.OppositeStartPos <> 0 AND #AUX.DDirection = 2)
               THEN
                   IF #DownDrill.AlreadyDrillLength <> 0 THEN
                       IF #DownDrill.AlreadyDrillLength > #DownDrill.SlabLength THEN
                           #DownDrill.OppositeStartPos := #DownDrill.SlabLength;
                       ELSE
                           #DownDrill.OppositeStartPos := #DownDrill.AlreadyDrillLength;
                       END_IF;
                   END_IF;
                   #DownDrill.PosNo := 0;
                   #DownDrill.AlreadyDrillLength := 0;
                   #DownDrill.gi_OffsetX := #DownDrill.AlreadyDrillWidth + #DownDrill.CurrentDrillWidth;
                   #DownDrill.AlreadyDrillWidth := #DownDrill.AlreadyDrillWidth + #DownDrill.CurrentDrillWidth;
                   IF #AUX.DDirection = 1 THEN
                       #AUX.DDirection := 2;
                       IF "DB720_KuKa_MainCtrl".CmdOut.gi_ToolTypeNo = 2 THEN
                           IF #DownDrill.OppositeStartPos + #DownDrill.CurrentDrillWidth / 2 > #DownDrill.SlabLength THEN
                               #DownDrill.OppositeStartPos := #DownDrill.OppositeStartPos - #DownDrill.CurrentDrillWidth / 2;
                           ELSE
                               #DownDrill.OppositeStartPos := #DownDrill.OppositeStartPos + #DownDrill.CurrentDrillWidth / 2;
                           END_IF;
                       END_IF;
                       IF "DB720_KuKa_MainCtrl".CmdOut.gi_ToolTypeNo = 13 THEN
                           IF "DB1900_Communication_PC".Para.DrillWidth = 65.0 THEN
                               #DownDrill.OppositeStartPos := 966.7;
                           END_IF;
                       END_IF;
                   ELSE
                       #AUX.DDirection := 1;
                       #DownDrill.gi_OffSetY := 0;
                       #DownDrill.OppositeStartPos := 0;
                   END_IF;
               ELSE
                   IF #AUX.DDirection = 1 THEN
                       #DownDrill.gi_OffSetY := #DownDrill.AlreadyDrillLength;
                   ELSE
                       #DownDrill.gi_OffSetY := #DownDrill.OppositeStartPos - #DownDrill.AlreadyDrillLength;
                   END_IF;
                   IF #DownDrill.CurrentDrillWidth <> #DownDrill.LastDrillWidth AND #DownDrill.PosNo <> 1 THEN
                       #DownDrill.AlreadyDrillWidth := #DownDrill.AlreadyDrillWidth + ABS(#DownDrill.CurrentDrillWidth / 2 - #DownDrill.LastDrillWidth / 2);
                       #DownDrill.gi_OffsetX := #DownDrill.AlreadyDrillWidth;
                       #DownDrill.LastDrillWidth := #DownDrill.CurrentDrillWidth;
                   END_IF;
               END_IF;
           ELSE
               "DB1900_Communication_PC".Send.PowerOff := TRUE;
               "DB1147_PromptStartNotPmt".Public.ChangeDownloadSlab := TRUE;
           END_IF;
       END_IF;
   END_IF;

   // ---------- 网络 8 ----------
   // 标题：当前水泥块已用完，请更换！
   // 含义：将 ("AutoMode_M" AND "DB1147_PromptStartNotPmt".Public.ChangeHorDrillSlab) OR ("AutoMode_M" AND "DB1147_PromptStartNotPmt".Public.ChangeHorVChiselSlab) OR ("AutoMode_M" AND "DB1147_PromptStartNotPmt".Public.ChangeDownloadSlab) 赋给 "DB1148_PromptBeeper".Public.ConcreteEnd
   "DB1148_PromptBeeper".Public.ConcreteEnd := ("AutoMode_M" AND "DB1147_PromptStartNotPmt".Public.ChangeHorDrillSlab) OR ("AutoMode_M" AND "DB1147_PromptStartNotPmt".Public.ChangeHorVChiselSlab) OR ("AutoMode_M" AND "DB1147_PromptStartNotPmt".Public.ChangeDownloadSlab);

   // ---------- 网络 9 ----------
   // （空白网络）
END_FUNCTION_BLOCK

// folder: 005_Component

FUNCTION_BLOCK "FB1080_Component"   // FB1080, SCL
{ S7_Optimized_Access := 'TRUE' }
// ============================================================
//  Block: FB1080_Component
//  ============================================================
//  编号：FB1080
//  原始语言：LAD（规则翻译为 SCL）
//  含义：******************************************************************************
//  ******************************************************************************
//  ******************************************************************************
//  ****************************   所有气缸的操作都在FB1081   **********************
//  ******************************************************************************
//  ******************************************************************************
//  ******************************************************************************
   VAR_INPUT
      ManMode : Bool;   // 输入参数
      AllMode : Bool;   // 输入参数
      EMMode : Bool;   // 输入参数
      ErrRst : Bool;   // 输入参数
      RobotEnble : Bool;   // 输入参数
      PromptStruct : Struct   // 输入参数
         Info : Struct   // 输入参数
            bit0 : Bool;   // 输入参数
            bit1 : Bool;   // 输入参数
            bit2 : Bool;   // 输入参数
            bit3 : Bool;   // 输入参数
            bit4 : Bool;   // 输入参数
            bit5 : Bool;   // 输入参数
            bit6 : Bool;   // 输入参数
            bit7 : Bool;   // 输入参数
            bit8 : Bool;   // 输入参数
            bit9 : Bool;   // 输入参数
            bit10 : Bool;   // 输入参数
            bit11 : Bool;   // 输入参数
            bit12 : Bool;   // 输入参数
            bit13 : Bool;   // 输入参数
            bit14 : Bool;   // 输入参数
            bit15 : Bool;   // 输入参数
            bit16 : Bool;   // 输入参数
            bit17 : Bool;   // 输入参数
            bit18 : Bool;   // 输入参数
            bit19 : Bool;   // 输入参数
            bit20 : Bool;   // 输入参数
            bit21 : Bool;   // 输入参数
            bit22 : Bool;   // 输入参数
            bit23 : Bool;   // 输入参数
            bit24 : Bool;   // 输入参数
            bit25 : Bool;   // 输入参数
            bit26 : Bool;   // 输入参数
            bit27 : Bool;   // 输入参数
            bit28 : Bool;   // 输入参数
            bit29 : Bool;   // 输入参数
            bit30 : Bool;   // 输入参数
            bit31 : Bool;   // 输入参数
         END_STRUCT;
         Err : Struct   // 输入参数
            bit0 : Bool;   // 输入参数
            bit1 : Bool;   // 输入参数
            bit2 : Bool;   // 输入参数
            bit3 : Bool;   // 输入参数
            bit4 : Bool;   // 输入参数
            bit5 : Bool;   // 输入参数
            bit6 : Bool;   // 输入参数
            bit7 : Bool;   // 输入参数
            bit8 : Bool;   // 输入参数
            bit9 : Bool;   // 输入参数
            bit10 : Bool;   // 输入参数
            bit11 : Bool;   // 输入参数
            bit12 : Bool;   // 输入参数
            bit13 : Bool;   // 输入参数
            bit14 : Bool;   // 输入参数
            bit15 : Bool;   // 输入参数
            bit16 : Bool;   // 输入参数
            bit17 : Bool;   // 输入参数
            bit18 : Bool;   // 输入参数
            bit19 : Bool;   // 输入参数
            bit20 : Bool;   // 输入参数
            bit21 : Bool;   // 输入参数
            bit22 : Bool;   // 输入参数
            bit23 : Bool;   // 输入参数
            bit24 : Bool;   // 输入参数
            bit25 : Bool;   // 输入参数
            bit26 : Bool;   // 输入参数
            bit27 : Bool;   // 输入参数
            bit28 : Bool;   // 输入参数
            bit29 : Bool;   // 输入参数
            bit30 : Bool;   // 输入参数
            bit31 : Bool;   // 输入参数
         END_STRUCT;
      END_STRUCT;
      IN : Bool;   // 输入参数
      TV : Time;   // 输入参数
      AlmEnable : Bool;   // 输入参数
      i_ID00 : Bool;   // 输入参数
      i_ID01 : Bool;   // 输入参数
      i_ID02 : Bool;   // 输入参数
      i_ID03 : Bool;   // 输入参数
      i_ID04 : Bool;   // 输入参数
      i_ID05 : Bool;   // 输入参数
      ParaR_FixIDCode : Byte;   // 输入参数
      Sys_Parameter_R_Gain : Real;   // 输入参数
      Sys_Parameter_R_Offset : Real;   // 输入参数
      IW_Analog : Int;   // 输入参数
      Type_Parameter_R_LimitMin : Real;   // 输入参数
      Type_Parameter_R_LimitMax : Real;   // 输入参数
      Sys_Parameter_R_AI_Gain : Real;   // 输入参数
      Sys_Parameter_R_AI_Offset : Real;   // 输入参数
      i_DoorOverRide : Bool;   // 输入参数
      i_AutoRunning : Bool;   // 输入参数
      i_OpenDoorPmt : Bool;   // 输入参数
   END_VAR
   VAR_OUTPUT
      PromptValue : Int;   // 输出参数
      Q : Bool;   // 输出参数
      Err : Bool;   // 输出参数
      QW_Analog_Out : Int;   // 输出参数
      o_DoorOverRideRelayOn : Bool;   // 输出参数
      o_DoorLockRelayON : Bool;   // 输出参数
      o_DoorOverRideLight : Bool;   // 输出参数
      o_PromptDoorOverRideStartIng : Bool;   // 输出参数
      o_PromptDoorOveRideStarted : Bool;   // 输出参数
      o_PromptDoorLockFail : Bool;   // 输出参数
   END_VAR
   VAR_IN_OUT
      Sys_Parameter_E_Gain : Real;   // 输入输出参数
      Sys_Parameter_E_Offset : Real;   // 输入输出参数
      Sys_Parameter_E_AI_Gain : Real;   // 输入输出参数
      Sys_Parameter_E_AI_Offset : Real;   // 输入输出参数
      IW : Int;   // 输入输出参数
      OUT_Offset : Real;   // 输入输出参数
      OUT_Gain : Real;   // 输入输出参数
   END_VAR
   VAR
      Robot : "FB5715_Kuka_General";   // 静态变量
      PowerFixtureID : "FB5003_FixtureID";   // 静态变量
      IOFixtureIID : "FB5003_FixtureID";   // 静态变量
      Analog_Out : "FB5007_Analog_Out_V3";   // 静态变量
      Press : "FB5006_Analog_IN_V4";   // 静态变量
      ClinyderPos : "FB5006_Analog_IN_V4";   // 静态变量
      SafetyDoor : "FB5002_SafetyDoorV1";   // 静态变量
      Analog_Out_1 : "FB5009_AnalOut";   // 静态变量
      Aux : Struct   // 静态变量
         Z08ExtPulse : Bool;   // 静态变量
         Pressure : Real;   // 静态变量
         PressureMid : Real;   // 静态变量
         Heart : IEC_TIMER;   // 静态变量
         HeartFalse : IEC_TIMER;   // 静态变量
      END_STRUCT;
      TP_Cmd : Word;   // 静态变量
      TP_Status : Word;   // 静态变量
      Cmd : Struct   // 静态变量
         Auto : Struct   // 静态变量
            ProgStart : Bool;   // 静态变量
            GoHome : Bool;   // 静态变量
            Stop : Bool;   // 静态变量
         END_STRUCT;
      END_STRUCT;
      CTRL_IN : Struct   // 静态变量
         ProgNo : Byte;   // 静态变量
         RobotSpeed : Byte;   // 静态变量
         InitParameter : Struct   // 静态变量
            HW_Addr : Hw_Io;   // 静态变量
            TimeOutSetValue : Time;   // 静态变量
            Td : Time;   // 静态变量
            sp : Array[0..3] of Real;   // 静态变量
         END_STRUCT;
      END_STRUCT;
      CTRL_OUT : Struct   // 静态变量
         ProgNo : Byte;   // 静态变量
         AppInfNo : Byte;   // 静态变量
         ErrorCode : Word;   // 静态变量
         LastCylceTime : Time;   // 静态变量
         sp : Array[1..16] of Byte;   // 静态变量
      END_STRUCT;
      Status : Struct   // 静态变量
         Busy : Bool;   // 静态变量
         OkToStart : Bool;   // 静态变量
         NotReadyV2 : Bool;   // 静态变量
         TaskDone : Bool;   // 静态变量
         TaskIO : Bool;   // 静态变量
         TaskNIO : Bool;   // 静态变量
         HomePos : Bool;   // 静态变量
         PromptValue : Int;   // 静态变量
      END_STRUCT;
      "Step" : Struct   // 静态变量
         Main : Int;   // 静态变量
      END_STRUCT;
      CmdMid : Struct   // 静态变量
         ProgStart : Bool;   // 静态变量
         GoHome : Bool;   // 静态变量
         Stop : Bool;   // 静态变量
      END_STRUCT;
      Bus_IN_Data : Struct   // 静态变量
         AlarmStop : Bool;   // 静态变量
         UserSaf : Bool;   // 静态变量
         Stopmess : Bool;   // 静态变量
         Alarm_Stop_Intern : Bool;   // 静态变量
         Pro_Act : Bool;   // 静态变量
         IN_home : Bool;   // 静态变量
         On_Path : Bool;   // 静态变量
         Robot_Rdy : Bool;   // 静态变量
         T1 : Bool;   // 静态变量
         T2 : Bool;   // 静态变量
         AUT : Bool;   // 静态变量
         EXT : Bool;   // 静态变量
         Peri_Rdy : Bool;   // 静态变量
         Rob_Stopped : Bool;   // 静态变量
         SP02 : Bool;   // 静态变量
         SP03 : Bool;   // 静态变量
         RecoveryActive : Bool;   // 静态变量
         CmdDone : Bool;   // 静态变量
         CmdRdy : Bool;   // 静态变量
         ProgReset : Bool;   // 静态变量
         SP04 : Byte;   // 静态变量
         Go_iCmd : Byte;   // 静态变量
         Go_iApplErrNo : Byte;   // 静态变量
         Go_iApplInfNo : Byte;   // 静态变量
         Gp330 : Byte;   // 静态变量
         UserDefineRobOut : Array[8..63] of Byte;   // 静态变量
      END_STRUCT;
      Bus_Out_Data : Struct   // 静态变量
         Move_Enable : Bool;   // 静态变量
         Ext_Start : Bool;   // 静态变量
         Conf_Mess : Bool;   // 静态变量
         Drives_On : Bool;   // 静态变量
         Drives_Off : Bool;   // 静态变量
         SP01 : Bool;   // 静态变量
         SP02 : Bool;   // 静态变量
         SP03 : Bool;   // 静态变量
         Recovery : Bool;   // 静态变量
         Ext_Stop : Bool;   // 静态变量
         AplFaultQuit : Bool;   // 静态变量
         CmdStart : Bool;   // 静态变量
         SP04 : Byte;   // 静态变量
         SP05 : Byte;   // 静态变量
         Gi_iCmd : Byte;   // 静态变量
         Gi_iRobotSpeed : Byte;   // 静态变量
         SP06 : Byte;   // 静态变量
         SP07 : Byte;   // 静态变量
         UserDefineRobIn : Array[8..63] of Byte;   // 静态变量
      END_STRUCT;
      Info_Err : Struct   // 静态变量
         InfoStruct : Struct   // 静态变量
            ModeOff : Bool;   // 静态变量
            OKToStart : Bool;   // 静态变量
            WaitUserCmdOff : Bool;   // 静态变量
            sp03 : Bool;   // 静态变量
            WaitBusyOff : Bool;   // 静态变量
            WaitIO_END : Bool;   // 静态变量
            WaitIO_Move : Bool;   // 静态变量
            WatiCmdRdy : Bool;   // 静态变量
            WaitChangeProg : Bool;   // 静态变量
            Sp11 : Bool;   // 静态变量
            Sp12 : Bool;   // 静态变量
            sp13 : Bool;   // 静态变量
            StartChangeProg : Bool;   // 静态变量
            DriversOn : Bool;   // 静态变量
            Ext_Start : Bool;   // 静态变量
            Recovery : Bool;   // 静态变量
            CmdStart : Bool;   // 静态变量
            CmdDone : Bool;   // 静态变量
            xx_5 : Bool;   // 静态变量
            xx_4 : Bool;   // 静态变量
            xx_3 : Bool;   // 静态变量
            xx : Bool;   // 静态变量
            xx_1 : Bool;   // 静态变量
            xx_2 : Bool;   // 静态变量
            xx_10 : Bool;   // 静态变量
            xx_11 : Bool;   // 静态变量
            xx_12 : Bool;   // 静态变量
            x : Bool;   // 静态变量
            xx_13 : Bool;   // 静态变量
            x_1 : Bool;   // 静态变量
            x_2 : Bool;   // 静态变量
            A37 : Bool;   // 静态变量
         END_STRUCT;
         ErrStruct : Struct   // 静态变量
            BusConnectErr : Bool;   // 静态变量
            EndOfTimeOut : Bool;   // 静态变量
            AlarmStopErr : Bool;   // 静态变量
            UserSafErr : Bool;   // 静态变量
            StopMessErr : Bool;   // 静态变量
            AlarmStopInternErr : Bool;   // 静态变量
            T1Mode : Bool;   // 静态变量
            T2Mode : Bool;   // 静态变量
            AutMode : Bool;   // 静态变量
            RobotNotRdy : Bool;   // 静态变量
            Sp12 : Bool;   // 静态变量
            sp37 : Bool;   // 静态变量
            sp36 : Bool;   // 静态变量
            sp35 : Bool;   // 静态变量
            sp34 : Bool;   // 静态变量
            sp33 : Bool;   // 静态变量
            sp31 : Bool;   // 静态变量
            xx_7 : Bool;   // 静态变量
            xx_6 : Bool;   // 静态变量
            xx_5 : Bool;   // 静态变量
            xx_4 : Bool;   // 静态变量
            xx : Bool;   // 静态变量
            xx_1 : Bool;   // 静态变量
            x : Bool;   // 静态变量
            x_1 : Bool;   // 静态变量
            x_2 : Bool;   // 静态变量
            x_3 : Bool;   // 静态变量
            x_4 : Bool;   // 静态变量
            x_5 : Bool;   // 静态变量
            x_6 : Bool;   // 静态变量
            E36 : Bool;   // 静态变量
            E37 : Bool;   // 静态变量
         END_STRUCT;
      END_STRUCT;
      FB_Prompt_Object : "FB1022_Prompt_ObjectV2";   // 静态变量
      Timer_TimeOut : "FB951_SDTimerV2";   // 静态变量
      TimdDrivers_Off : "FB951_SDTimerV2";   // 静态变量
      Stack : Struct   // 静态变量
         Index : Int;   // 静态变量
         "Step" : Array[0..9] of Int;   // 静态变量
         sp : Array[0..1] of Int;   // 静态变量
      END_STRUCT;
      lastAddr : Int;   // 静态变量
      CycleTime : Int;   // 静态变量
      PromptValueBake : Int;   // 静态变量
      ShiftBake : Int;   // 静态变量
      StartTime : Time;   // 静态变量
      ET : Time;   // 静态变量
      IN_EDGE : Bool;   // 静态变量
      TP_CurFixtureID : Byte;   // 静态变量
      sp : Int;   // 静态变量
      TP_DoorInsert : Array[1..8] of Bool;   // 静态变量
      TP_DoorUnLock : Array[1..8] of Bool;   // 静态变量
      Confirm : Bool;   // 静态变量
      PT : Time;   // 静态变量
   END_VAR
   VAR_TEMP
      OverAllPmt : Bool;   // 临时变量
      Ret : Int;   // 临时变量
   END_VAR
BEGIN

   // ---------- 网络 1 ----------
   // 标题：所有模式
   // 含义：将 "ICurtainsOK" AND NOT (#SafetyDoor.i_DoorOverRide) 赋给 #OverAllPmt
   #OverAllPmt := "ICurtainsOK" AND NOT (#SafetyDoor.i_DoorOverRide);
   // 含义：当 "ICurtainsOK" 为 TRUE 时置位 "QCurtainRst"，否则复位（触点→线圈）
   IF "ICurtainsOK" THEN
       "QCurtainRst" := TRUE;
   ELSE
       "QCurtainRst" := FALSE;
   END_IF;
   // 含义：将 (NOT ("IAirPressOK") OR NOT ("ICurtainsOK")) AND "DB1000_StdSignal".RectWave.Wave05 赋给 "QCurtainLight"
   "QCurtainLight" := (NOT ("IAirPressOK") OR NOT ("ICurtainsOK")) AND "DB1000_StdSignal".RectWave.Wave05;
   // 含义：当 "DB1900_Communication_PC".Recv.Heart 为 TRUE 时置位 "DB1900_Communication_PC".Send.Heart，否则复位（触点→线圈）
   IF "DB1900_Communication_PC".Recv.Heart THEN
       "DB1900_Communication_PC".Send.Heart := TRUE;
   ELSE
       "DB1900_Communication_PC".Send.Heart := FALSE;
   END_IF;
   // 含义：调用计数器实例 #Aux.Heart.TON（上升沿计数，当前值写入 CV）
   #Aux.Heart.TON(IN := "DB1900_Communication_PC".Recv.Heart,
                  PT := T#10S);
   // 含义：条件 "DB1900_Communication_PC".Recv.Heart AND "ErrRst_M" 成立时，将 FALSE 传送到 "DB1147_PromptStartNotPmt".Public.PcCommErr
   IF "DB1900_Communication_PC".Recv.Heart AND "ErrRst_M" THEN
       "DB1147_PromptStartNotPmt".Public.PcCommErr := FALSE;
   END_IF;
   // 含义：调用计数器实例 #Aux.HeartFalse.TON（上升沿计数，当前值写入 CV）
   #Aux.HeartFalse.TON(IN := NOT ("DB1900_Communication_PC".Recv.Heart),
                       PT := T#10S);
   // 含义：条件 #Aux.Heart.Q OR #Aux.HeartFalse.Q 成立时，将 TRUE 传送到 "DB1147_PromptStartNotPmt".Public.PcCommErr
   IF #Aux.Heart.Q OR #Aux.HeartFalse.Q THEN
       "DB1147_PromptStartNotPmt".Public.PcCommErr := TRUE;
   END_IF;
   // 含义：条件 #Aux.Heart.Q OR #Aux.HeartFalse.Q 成立时，将 TRUE 传送到 "DB1900_Communication_PC".Send.PowerOff
   IF #Aux.Heart.Q OR #Aux.HeartFalse.Q THEN
       "DB1900_Communication_PC".Send.PowerOff := TRUE;
   END_IF;
   // 含义：条件 #Aux.Heart.Q OR #Aux.HeartFalse.Q 成立时，将 TRUE 传送到 #Robot.Cmd.Auto.Stop
   IF #Aux.Heart.Q OR #Aux.HeartFalse.Q THEN
       #Robot.Cmd.Auto.Stop := TRUE;
   END_IF;
   // 含义：条件 NOT ("AllMode_M") 成立时，将 TRUE 传送到 #Robot.Cmd.Auto.Stop
   IF NOT ("AllMode_M") THEN
       #Robot.Cmd.Auto.Stop := TRUE;
   END_IF;
   // 含义：条件 NOT ("AllMode_M") 成立时，将 TRUE 传送到 "DB1081_ValveCall".ST01.Z05.RetAuto
   IF NOT ("AllMode_M") THEN
       "DB1081_ValveCall".ST01.Z05.RetAuto := TRUE;
   END_IF;
   // 含义：条件 NOT ("EMMode_M") AND NOT (#Aux.Z08ExtPulse) 成立时，将 TRUE 传送到 "DB1081_ValveCall".ST01.Z08.ExtAuto
   IF NOT ("EMMode_M") AND NOT (#Aux.Z08ExtPulse) THEN
       "DB1081_ValveCall".ST01.Z08.ExtAuto := TRUE;
   END_IF;
   // 含义：条件 NOT ("EMMode_M") AND NOT (#Aux.Z08ExtPulse) 成立时，将 0.4 传送到 #Aux.Pressure
   IF NOT ("EMMode_M") AND NOT (#Aux.Z08ExtPulse) THEN
       #Aux.Pressure := 0.4;
   END_IF;
   // 含义：当 NOT ("EMMode_M") 为 TRUE 时置位 #Aux.Z08ExtPulse，否则复位（触点→线圈）
   IF NOT ("EMMode_M") THEN
       #Aux.Z08ExtPulse := TRUE;
   ELSE
       #Aux.Z08ExtPulse := FALSE;
   END_IF;

   // ---------- 网络 2 ----------
   // 标题：标准动作的控制
   // 注释：******************************************************************************
   // ******************************************************************************
   // ******************************************************************************
   // ****************************   所有气缸的操作都在FB1081   **********************
   // ******************************************************************************
   // ******************************************************************************
   // ******************************************************************************
   // 含义：调用块/实例 "DB1081_ValveCall"
   "DB1081_ValveCall"();

   // ---------- 网络 3 ----------
   // 标题：SafeDoor
   // 含义：调用定时器实例 #SafetyDoor
   #SafetyDoor(i_DoorOverRide := "IDoorOverRide",
               i_AutoRunning := "ASMMode_M",
               i_OpenDoorPmt := "IMan",
               EMMode := "EMMode_M",
               o_DoorLockRelayON => "QDoorClose",
               o_DoorOverRideLight => "QSpairMode",
               o_PromptDoorOveRideStarted => "DB1147_PromptStartNotPmt".Public.DoorOveRideStarted);

   // ---------- 网络 4 ----------
   // 标题：Robot
   // 含义：条件 NOT ("AllMode_M") 成立时，将 "AG1521Kuka_Big~512_digital_in-_and_outputs_1" 传送到 #Robot.CTRL_IN.InitParameter.HW_Addr
   IF NOT ("AllMode_M") THEN
       #Robot.CTRL_IN.InitParameter.HW_Addr := "AG1521Kuka_Big~512_digital_in-_and_outputs_1";
   END_IF;
   // 含义：当 #OverAllPmt 为 TRUE 时置位 #Robot.RobotEnble，否则复位（触点→线圈）
   IF #OverAllPmt THEN
       #Robot.RobotEnble := TRUE;
   ELSE
       #Robot.RobotEnble := FALSE;
   END_IF;
   // 含义：将 "AllMode_M" AND #Robot.Status.NotReadyV2 赋给 "DB1148_PromptBeeper".Public.RobotNotReady
   "DB1148_PromptBeeper".Public.RobotNotReady := "AllMode_M" AND #Robot.Status.NotReadyV2;
   // 含义：条件 "AllMode_M" AND #Robot.Status.NotReadyV2 成立时，将 TRUE 传送到 "DB1900_Communication_PC".Send.PowerOff
   IF "AllMode_M" AND #Robot.Status.NotReadyV2 THEN
       "DB1900_Communication_PC".Send.PowerOff := TRUE;
   END_IF;
   // 含义：调用块/实例 "DB720_KuKa_MainCtrl"
   "DB720_KuKa_MainCtrl"();
   // 含义：调用块/实例 #Robot，参数：ManMode := "ManMode_M", AllMode := "AllMode_M", EMMode := "EMMode_M", ErrRst := "ErrRst_M"
   #Robot(ManMode := "ManMode_M",
          AllMode := "AllMode_M",
          EMMode := "EMMode_M",
          ErrRst := "ErrRst_M");

   // ---------- 网络 5 ----------
   // 标题：钻孔数据计算
   // 含义：调用块/实例 "DB1910_DrillData"
   "DB1910_DrillData"();

   // ---------- 网络 6 ----------
   // 标题：夹具编码
   // 含义：调用块/实例 #PowerFixtureID，参数：i_ID00 := "IFixtureCode01", i_ID01 := "IFixtureCode02", i_ID02 := "IFixtureCode03", ParaR_FixIDCode := "DB1900_Communication_PC".Para.PowerFixtureNo
   #PowerFixtureID(i_ID00 := "IFixtureCode01",
                   i_ID01 := "IFixtureCode02",
                   i_ID02 := "IFixtureCode03",
                   ParaR_FixIDCode := "DB1900_Communication_PC".Para.PowerFixtureNo);
   // 含义：调用块/实例 #IOFixtureIID，参数：i_ID00 := "IFixtureIOCode01", i_ID01 := "IFixtureIOCode02", i_ID02 := "IFixtureIOCode03", ParaR_FixIDCode := "DB1900_Communication_PC".Para.IOFixtureNo
   #IOFixtureIID(i_ID00 := "IFixtureIOCode01",
                 i_ID01 := "IFixtureIOCode02",
                 i_ID02 := "IFixtureIOCode03",
                 ParaR_FixIDCode := "DB1900_Communication_PC".Para.IOFixtureNo);

   // ---------- 网络 7 ----------
   // 标题：压力
   // 含义：调用定时器实例 #Press
   #Press(ManMode := "ManMode_M",
          IW_Analog := "IW10",
          Sys_Parameter_R_AI_Gain := "DB1010_Parameter".SystemParaR.Other.IN_Gain,
          Sys_Parameter_R_AI_Offset := "DB1010_Parameter".SystemParaR.Other.IN_Offset,
          Sys_Parameter_E_AI_Gain := "DB1010_Parameter".SystemParaE.Other.IN_Gain,
          Sys_Parameter_E_AI_Offset := "DB1010_Parameter".SystemParaE.Other.IN_Offset);

   // ---------- 网络 8 ----------
   // 标题：推力位置
   // 含义：调用定时器实例 #ClinyderPos
   #ClinyderPos(ManMode := "ManMode_M",
                IW_Analog := "IW12",
                Sys_Parameter_R_AI_Gain := "DB1010_Parameter".SystemParaR.Other.IN_Gain_1,
                Sys_Parameter_R_AI_Offset := "DB1010_Parameter".SystemParaR.Other.IN_Offset_1,
                Sys_Parameter_E_AI_Gain := "DB1010_Parameter".SystemParaE.Other.IN_Gain_1,
                Sys_Parameter_E_AI_Offset := "DB1010_Parameter".SystemParaE.Other.IN_Offset_1);

   // ---------- 网络 9 ----------
   // 含义：调用定时器实例 #Analog_Out_1
   #Analog_Out_1(IW := "QW10",
                 OUT_Offset := "DB1010_Parameter".SystemParaE.Other.OUT_Offset,
                 OUT_Gain := "DB1010_Parameter".SystemParaE.Other.OUT_Gain);
   // 含义：条件 (#Aux.Pressure >= 0.6) 成立时，将 0.6 传送到 #Aux.Pressure
   IF (#Aux.Pressure >= 0.6) THEN
       #Aux.Pressure := 0.6;
   END_IF;
   // 含义：将 (#Aux.Pressure - "DB1010_Parameter".SystemParaR.Other.OUT_Offset) 赋给 #Aux.PressureMid
   #Aux.PressureMid := (#Aux.Pressure - "DB1010_Parameter".SystemParaR.Other.OUT_Offset);
   // 含义：将 (#Aux.PressureMid / "DB1010_Parameter".SystemParaR.Other.OUT_Gain) 赋给 "QW10"
   "QW10" := (#Aux.PressureMid / "DB1010_Parameter".SystemParaR.Other.OUT_Gain);

   // ---------- 网络 10 ----------
   // 含义：调用块/实例 FC1900_Communication_PC
   "FC1900_Communication_PC"();

   // ---------- 网络 11 ----------
   // 标题：报警信息
   // 含义：条件 "AllMode_M" 成立时，将 0 传送到 "DB1900_Communication_PC".Send.Beer_info
   IF "AllMode_M" THEN
       "DB1900_Communication_PC".Send.Beer_info := 0;
   END_IF;
   // 含义：条件 "AllMode_M" AND "DB1148_PromptBeeper".Public.CurrentLowTimeOut 成立时，将 2029 传送到 "DB1900_Communication_PC".Send.Beer_info
   IF "AllMode_M" AND "DB1148_PromptBeeper".Public.CurrentLowTimeOut THEN
       "DB1900_Communication_PC".Send.Beer_info := 2029;
   END_IF;
   // 含义：条件 "AllMode_M" AND "DB1148_PromptBeeper".Public.DrillDepthErr 成立时，将 2030 传送到 "DB1900_Communication_PC".Send.Beer_info
   IF "AllMode_M" AND "DB1148_PromptBeeper".Public.DrillDepthErr THEN
       "DB1900_Communication_PC".Send.Beer_info := 2030;
   END_IF;
   // 含义：条件 "AllMode_M" AND "DB1148_PromptBeeper".Public.DrillTimeOut 成立时，将 2005 传送到 "DB1900_Communication_PC".Send.Beer_info
   IF "AllMode_M" AND "DB1148_PromptBeeper".Public.DrillTimeOut THEN
       "DB1900_Communication_PC".Send.Beer_info := 2005;
   END_IF;

   // ---------- 网络 12 ----------
   // 含义：调用块/实例 "DB2008_CoolingFan[DB2008]"
   "DB2008_CoolingFan[DB2008]"();

   // ---------- 网络 13 ----------
   // （空白网络）
END_FUNCTION_BLOCK

FUNCTION_BLOCK "FB5003_FixtureID"   // FB5003, SCL
{ S7_Optimized_Access := 'TRUE' }
// ============================================================
//  Block: FB5003_FixtureID
//  ============================================================
//  编号：FB5003
//  原始语言：LAD（规则翻译为 SCL）
//  含义：由 LAD/FBD 网络折叠生成的等效 SCL，导入前请人工复核
   VAR_INPUT
      AlmEnable : Bool := TRUE;   // 输入参数
      i_ID00 : Bool;   // 输入参数
      i_ID01 : Bool;   // 输入参数
      i_ID02 : Bool;   // 输入参数
      i_ID03 : Bool;   // 输入参数
      i_ID04 : Bool;   // 输入参数
      i_ID05 : Bool;   // 输入参数
      ParaR_FixIDCode : Byte;   // 参数设置的夹具编码
   END_VAR
   VAR_OUTPUT
      Err : Bool;   // 夹具编码不匹配，请更换夹具！
   END_VAR
   VAR
      TP_CurFixtureID : Byte;   // 用于触摸屏显示当前夹具编码状态
      sp : Int;   // 静态变量
      LastAddr : Int := 8;   // 静态变量
   END_VAR
BEGIN

   // ---------- 网络 1 ----------
   // 标题：转存当前实际的夹具编码
   // 含义：当 #i_ID00 为 TRUE 时置位 #TP_CurFixtureID，否则复位（触点→线圈）
   #TP_CurFixtureID.%X0 := #i_ID00;
   #TP_CurFixtureID.%X1 := #i_ID01;
   #TP_CurFixtureID.%X2 := #i_ID02;
   #TP_CurFixtureID.%X3 := #i_ID03;
   #TP_CurFixtureID.%X4 := #i_ID04;
   #TP_CurFixtureID.%X5 := #i_ID05;
   #TP_CurFixtureID.%X6 := FALSE;
   #TP_CurFixtureID.%X7 := FALSE;

   // ---------- 网络 2 ----------
   // 标题：对比给出报警信息
   // 含义：将 (#ParaR_FixIDCode <> #TP_CurFixtureID) AND #AlmEnable 赋给 #Err
   #Err := (#ParaR_FixIDCode <> #TP_CurFixtureID) AND #AlmEnable;

   // ---------- 网络 3 ----------
   // （空白网络）
END_FUNCTION_BLOCK

FUNCTION_BLOCK "FB5006_Analog_IN_V4"   // FB5006, SCL
{ S7_Optimized_Access := 'TRUE' }
// ============================================================
//  Block: FB5006_Analog_IN_V4
//  ============================================================
//  编号：FB5006
//  原始语言：SCL（规则翻译为 SCL）
//  含义：由 LAD/FBD 网络折叠生成的等效 SCL，导入前请人工复核
   VAR_INPUT
      ManMode : Bool := TRUE;   // 手动模式
      IW_Analog : Int;   // 输入模拟量数值，来自AIW
      Type_Parameter_R_LimitMin : Real;   // 对比用的最小值，来自参数
      Type_Parameter_R_LimitMax : Real;   // 对比用的最大值，来自参数
      Sys_Parameter_R_AI_Gain : Real := 12.58;   // 来自运行区参数（800~1000）
      Sys_Parameter_R_AI_Offset : Real;   // 来自运行区参数
   END_VAR
   VAR_IN_OUT
      Sys_Parameter_E_AI_Gain : Real;   // 到编辑区参数
      Sys_Parameter_E_AI_Offset : Real;   // 到编辑区参数
   END_VAR
   VAR
      TP_Cmd : Word;   // 静态变量
      Cmd : Struct   // 静态变量
         Man : Struct   // 静态变量
            SetToPreSetValue : Bool;   // 根据期望值,计算增益;
            Record_ActualAI_1 : Bool;   // 记录两点校验的模拟量1
            Record_ActualAI_2 : Bool;   // 记录两点校验的模拟量2
            Calculate : Bool;   // 计算线性增益及偏置
         END_STRUCT;
         Auto : Struct   // 静态变量
            ClearCompareResult : Bool;   // 清除前次的对比输出结果
            ClearRecordCounter : Bool;   // 清除记录值的序号，同时清除对比输出结果
            TrigerCompare : Bool;   // 触发对比
         END_STRUCT;
      END_STRUCT;
      AtCmd : Struct   // 静态变量
         Man : Word;   // 静态变量
         Auto : Word;   // 静态变量
      END_STRUCT;
      Ctrl_IN : Struct   // 静态变量
         TP_AI_Gain : Real;   // 计算的增益
         TP_AI_OffSet : Real;   // 计算的偏置（补偿量）
         TP_PreSetValue : Real;   // 期望的预定义值，来自屏幕
         TP_ActualAI_1 : Real;   // 2点标定模拟量值1
         TP_ActualAI_2 : Real;   // 2点标定模拟量值2
         TP_ActualAI_Value1 : Real;   // 2点标定实际值1
         TP_ActualAI_Value2 : Real;   // 2点标定实际值2
         sp : Array[1..18] of Byte;   // 静态变量
      END_STRUCT;
      Ctrl_Out : Struct   // 静态变量
         Cur_Val_Out : Real;   // 当前值输出,可以用于屏幕显示
         TrigerValue : Real;   // 最近一次对比的记录值
         TrigerTPColorStatus : Int;   // 最近一次对比的结果输出,1:Less, 2: OK, 4: More
         TrigerValue_Array : Array[1..10] of Real;   // 对比值
         TrigerTPColorStatus_Array : Array[1..10] of Int;   // 1:Less, 2: OK, 4: More
         TrigerCounter : Int := 1;   // 静态变量
      END_STRUCT;
      Status : Struct   // 静态变量
         Low : Bool;   // 请求后判断的状态
         In : Bool;   // 请求后判断的状态
         High : Bool;   // 请求后判断的状态
         xxxxsp1 : Byte;   // 静态变量
         Low_Realtime : Bool;   // 实时值偏低
         In_Realtime : Bool;   // 实时值在范围内
         High_Realtime : Bool;   // 实时值偏大
         TrigerCompare_Done : Bool;   // 对比完成,数据已经更新
         Clear_Done : Bool;   // 清除完成
      END_STRUCT;
      AtStatus : Struct   // 静态变量
         CompareStatus : Byte;   // 静态变量
      END_STRUCT;
      Aux : Struct   // 静态变量
         AI_RealRawValue : Real;   // 取整为1
         AI_LinearValue : Real;   // 乘以增益后;
         Max_Anlog_Value_Real : Real := 27648.0;   // 静态变量
         sp : Array[1..30] of Byte;   // 静态变量
      END_STRUCT;
      LastAddr : Int := 198;   // 静态变量
   END_VAR
BEGIN
END_FUNCTION_BLOCK

FUNCTION_BLOCK "FB5007_Analog_Out_V3"   // FB5007, SCL
{ S7_Optimized_Access := 'TRUE' }
// ============================================================
//  Block: FB5007_Analog_Out_V3
//  ============================================================
//  编号：FB5007
//  原始语言：SCL（规则翻译为 SCL）
//  含义：由 LAD/FBD 网络折叠生成的等效 SCL，导入前请人工复核
   VAR_INPUT
      ManMode : Bool := TRUE;   // 手动模式
      Sys_Parameter_R_Gain : Real;   // 来自运行区参数
      Sys_Parameter_R_Offset : Real;   // 来自运行区参数
   END_VAR
   VAR_OUTPUT
      QW_Analog_Out : Int;   // 对应模拟量输出
   END_VAR
   VAR_IN_OUT
      Sys_Parameter_E_Gain : Real;   // 到编辑区参数
      Sys_Parameter_E_Offset : Real;   // 到编辑区参数
   END_VAR
   VAR
      TP_Cmd : Word;   // 静态变量
      Cmd : Struct   // 静态变量
         Man : Struct   // 静态变量
            SetToPreSetValue : Bool;   // 计算偏置值
            Record_ActualAnalog_1 : Bool;   // 静态变量
            Record_ActualAnalog_2 : Bool;   // 静态变量
            Calculate : Bool;   // 静态变量
         END_STRUCT;
      END_STRUCT;
      AtCmd : Struct   // 静态变量
         Man : Word;   // 静态变量
      END_STRUCT;
      Ctrl_IN : Struct   // 静态变量
         TP_Gain : Real;   // （工程单位）增益
         TP_Offset : Real;   // （工程单位）偏置
         TP_PresetValue : Real;   // （工程单位）预置值
         TP_ActualAO_1 : Real;   // 归一后的2点标定示教模拟量值_1
         TP_ActualAO_2 : Real;   // 归一后的2点标定示教模拟量值_2
         TP_ActualAO_Value1 : Real;   // （工程单位）2点标定示教值_1
         TP_ActualAO_Value2 : Real;   // （工程单位）2点标定示教值_2
         Target : Real;   // （工程单位）用于设定目标值
         Max_Anlog_Value_Real : Real := 27648.0;   // 静态变量
      END_STRUCT;
      Aux : Struct   // 静态变量
         Analog_Out_Real : Real;   // 取整为1
         SetToPreSetValuePulse : Bool;   // 静态变量
         Sp : Array[0..31] of Byte;   // 静态变量
      END_STRUCT;
      LastAddr : Int := 98;   // 静态变量
   END_VAR
BEGIN
END_FUNCTION_BLOCK

FUNCTION_BLOCK "FB5009_AnalOut"   // FB5009, SCL
{ S7_Optimized_Access := 'TRUE' }
// ============================================================
//  Block: FB5009_AnalOut
//  ============================================================
//  编号：FB5009
//  原始语言：LAD（规则翻译为 SCL）
//  含义：由 LAD/FBD 网络折叠生成的等效 SCL，导入前请人工复核
   VAR_IN_OUT
      IW : Int;   // 输入输出参数
      OUT_Offset : Real;   // 输入输出参数
      OUT_Gain : Real;   // 输入输出参数
   END_VAR
   VAR
      Confirm : Bool;   // 静态变量
      Ctrl_IN : Struct   // 静态变量
         TP_ActualAI_1 : Real;   // 2点标定模拟量值1
         TP_ActualAI_2 : Real;   // 2点标定模拟量值2
         TP_ActualAI_Value1 : Real;   // 2点标定实际值1
         TP_ActualAI_Value2 : Real;   // 2点标定实际值2
      END_STRUCT;
      Ctrl_Out : Struct   // 静态变量
         k : Real;   // 静态变量
         "b" : Real;   // 静态变量
         Pressure : Real;   // 静态变量
      END_STRUCT;
      Cmd : Struct   // 静态变量
         Read1 : Bool;   // 静态变量
         Read2 : Bool;   // 静态变量
      END_STRUCT;
   END_VAR
BEGIN

   // ---------- 网络 1 ----------
   // 含义：本网络为 StructuredText（SCL）原文重建，非 LAD 折叠
   #Ctrl_Out.b := (#Ctrl_IN.TP_ActualAI_Value2 * #Ctrl_IN.TP_ActualAI_1 - #Ctrl_IN.TP_ActualAI_Value1 * #Ctrl_IN.TP_ActualAI_2) / (#Ctrl_IN.TP_ActualAI_1 - #Ctrl_IN.TP_ActualAI_2);
   #Ctrl_Out.k := (#Ctrl_IN.TP_ActualAI_Value1 - #Ctrl_Out.b) / #Ctrl_IN.TP_ActualAI_1;

   // ---------- 网络 2 ----------
   // 含义：将 #IW; (* Convert → Real *) END_IF 赋给 IF #Cmd.Read1 THEN #Ctrl_IN.TP_ActualAI_1
   IF #Cmd.Read1 THEN
       #Ctrl_IN.TP_ActualAI_1 := #IW; (* Convert → Real *)
   END_IF;
   // 含义：将 #IW; (* Convert → Real *) END_IF 赋给 IF #Cmd.Read2 THEN #Ctrl_IN.TP_ActualAI_2
   IF #Cmd.Read2 THEN
       #Ctrl_IN.TP_ActualAI_2 := #IW; (* Convert → Real *)
   END_IF;

   // ---------- 网络 3 ----------
   // 含义：本网络为 StructuredText（SCL）原文重建，非 LAD 折叠
   IF #Confirm
   THEN
       #OUT_Offset := #Ctrl_Out.b;
       #OUT_Gain := #Ctrl_Out.k;
   END_IF;
   #Ctrl_Out.Pressure := #Ctrl_Out.k * #IW + #Ctrl_Out.b;

   // ---------- 网络 4 ----------
   // （空白网络）
END_FUNCTION_BLOCK

FUNCTION_BLOCK "FB5019_stringSegment"   // FB5019, SCL
{ S7_Optimized_Access := 'TRUE' }
// ============================================================
//  Block: FB5019_stringSegment
//  ============================================================
//  编号：FB5019
//  原始语言：SCL（规则翻译为 SCL）
//  含义：由 LAD/FBD 网络折叠生成的等效 SCL，导入前请人工复核
   VAR
      Ctrl_In : Struct   // 静态变量
         srcResultStr : String := 'abc,eft,aaa,aaa';   // 字符串,例如'abc,eft,aaa,aaa'
         SepeartorString : String[1] := ',';   // 分隔符，例如','
      END_STRUCT;
      Ctrl_OUT : Struct   // 静态变量
         SegNum : Int;   // 表示找到的分隔符数量
         str_Segment : Array[0..19] of String[18];   // 静态变量
      END_STRUCT;
      Aux : Struct   // 静态变量
         sp : Array[0..35] of Byte;   // 静态变量
      END_STRUCT;
      LastAddr : Int := 698;   // 静态变量
   END_VAR
BEGIN
END_FUNCTION_BLOCK

FUNCTION_BLOCK "FB5020_TypeConvert_4ByteDWORD_Real"   // FB5020, SCL
{ S7_Optimized_Access := 'TRUE' }
// ============================================================
//  Block: FB5020_TypeConvert_4ByteDWORD_Real
//  ============================================================
//  编号：FB5020
//  原始语言：SCL（规则翻译为 SCL）
//  含义：由 LAD/FBD 网络折叠生成的等效 SCL，导入前请人工复核
   VAR_INPUT
      DataType : Byte;   // 2-> int8; 3-> Int16; 4->Int32; 5,41-> U8, 6,42-> U16,7,43-> U32,8:Real
      Dword_DataIn : DWord;   // 待转换的值
      AtInt : Int;   // 3
      AtDint : DInt;   // 4
      AtReal : Real;   // 8
      AtByte : Byte;   // 5,41
      AtWord : Word;   // 6,42
      AtDword : DWord;   // 7,43
   END_VAR
   VAR_OUTPUT
      Real_DataOut : Real;   // 输出参数
      ErrCode : Int;   // 输出参数
      DataTypeError : Bool;   // 数据类型有误
   END_VAR
BEGIN
END_FUNCTION_BLOCK

FUNCTION_BLOCK "FB5021_TypeConvert_Real_4ByteDWord"   // FB5021, SCL
{ S7_Optimized_Access := 'TRUE' }
// ============================================================
//  Block: FB5021_TypeConvert_Real_4ByteDWord
//  ============================================================
//  编号：FB5021
//  原始语言：SCL（规则翻译为 SCL）
//  含义：由 LAD/FBD 网络折叠生成的等效 SCL，导入前请人工复核
   VAR_INPUT
      DataType : Byte;   // 2-> int8; 3-> Int16; 4->Int32; 5,41-> U8, 6,42-> U16,7,43-> U32,8:Real
      Real_DataIn : Real;   // 待转换的值
   END_VAR
   VAR_OUTPUT
      DWord_DataOut : DWord;   // 输出参数
      AtInt_DWord_ToSend : Int;   // 3
      AtDint_DWord_ToSend : DInt;   // 4
      AtReal_DWord_ToSend : Real;   // 8
      AtByte_DWord_ToSend : Byte;   // 5,41
      AtWord_DWord_ToSend : Word;   // 6,42
      AtDword_DWord_ToSend : DWord;   // 7,43
      DataTypeError : Bool;   // 数据类型有误
   END_VAR
BEGIN
END_FUNCTION_BLOCK

FUNCTION_BLOCK "FB5699_RandomDemoTest"   // FB5699, SCL
{ S7_Optimized_Access := 'TRUE' }
// ============================================================
//  Block: FB5699_RandomDemoTest
//  ============================================================
//  编号：FB5699
//  原始语言：LAD（规则翻译为 SCL）
//  含义：//*************************************************************************
//  //*********************上海克来机电自动化工程股份有限公司***********************
//  //***********************               V2017.02.15          ******************************
//  //**********************             功能块快速测试用         *****************************
//  //**********************                  乱序随机测试            *****************************
//  //**************************************************************************
//  First created on 2017.02.15；
   VAR_INPUT
      ManMode : Bool;   // 手动模式
      AllMode : Bool;   // 所有模式
      EMMode : Bool;   // 紧急停止模式
      ErrRst : Bool;   // 故障复位
      Pulse_En : Bool;   // 输入参数
      PromptSourceDW : DWord;   // 输入参数
      TV : Time;   // 输入参数
   END_VAR
   VAR_OUTPUT
      PromptValue : Int;   // 输出参数
   END_VAR
   VAR_IN_OUT
      Servo_Cmd : Struct   // 输入输出参数
         Man : Struct   // 输入输出参数
            StartHoming : Bool;   // Starts Homing Task
            StartTask : Bool;   // Starts Positioning Task
            TorqueCtrl_FixedStop : Bool;   // Starts Torque Control mode
            JogPos : Bool;   // Jogging positive direction
            JogNeg : Bool;   // Jogging negaitive direction
            HomeToWorkPos : Bool;   // Starts Work HomePosition
            StartTraversingBlock : Bool;   // Start Traversing block
            ServoOff_And_BrakeRelease : Bool;   // Servo and Brake release
            ParaWrite : Bool;   // Request parameter value (array, double word)
            ParaRead : Bool;   // Modify parameter value (array, double word)
            SetTLM : Bool;   // Set torqueLimit
            ResetTLM : Bool;   // ResetTorqueLimit
            StartTask_TLM : Bool;   // Starts Positioning Task with torque limited!
         END_STRUCT;
         Auto : Struct   // 输入输出参数
            StartHoming : Bool;   // Starts Homing Task
            StartTask : Bool;   // Starts Positioning Task
            TorqueCtrl_FixedStop : Bool;   // Starts Torque Control mode
            JogPos : Bool;   // Jogging positive direction
            JogNeg : Bool;   // Jogging negaitive direction
            HomeToWorkPos : Bool;   // Starts Work HomePosition
            StartTraversingBlock : Bool;   // Start Traversing block
            ServoOff_And_BrakeRelease : Bool;   // 关闭使能
            ParaWrite : Bool;   // Request parameter value (array, double word)
            ParaRead : Bool;   // Modify parameter value (array, double word)
            SetTLM : Bool;   // Set torqueLimit
            ResetTLM : Bool;   // ResetTorqueLimit
            StartTask_TLM : Bool;   // Starts Positioning Task with torque limited!
            Halt : Bool;   // Halt current command
            Stop : Bool;   // Stop Current command and output result TaskNIO
            ServoOff2 : Bool;   // ServoOff and no fault occur
         END_STRUCT;
      END_STRUCT;
      Servo_CTRL_IN : Struct   // 输入输出参数
         SetValueVelocity : Real;   // Setvalue Velocity %(Directmode/Positionmode)
         SetValuePosition : Real;   // SetValue Position (Directmode/Positioncontrol)
         SetWorkHomePos : Real;   // WorkHomePos
         SetValueTorque : Real;   // SetValueTorque_P2622
         TraversingBlockNO : Byte;   // Traversing block no. NO.0 is dedicated for fixed stop mode
         TraversingBlockCycleNO : DInt;   // Traversing Block 循环次数
         PNU : Int;   // the parameter number
         SubIndex : Byte;   // Addresses an element of an array parameter (sub-parameter number).
         ParameterValue_DataCom : Real;   // Value of the parameter to be write to Festo controller
         TrackingModeActive : Bool;   // user should keep this bit ON。
         EnTorqueLimited : Bool;   // Enanble torque limited with the coming motion
         ResetTLM_AfterTorqueCtrl : Bool;   // 执行完扭矩模式后，是否关闭扭矩模式！
         ModularEnable : Bool;   // whether enable Modular,是否开启模态轴
         InitParameter : Struct   // 输入输出参数
            InPosTolerance : Real;   // 默认--到位置范围精度*Lead
            Lead : Real;   // *_导程，即：p29247, set the length per revolution
            MaxRotationSpeedAfterGearBox : Real;   // 减速箱后的最大转速,例如额定3000rpm=50rps, 选择10的减速比,则最大转速50/10=5.0
            Min_SetValuePosition : Real;   // 负向运动的最小位置
            Max_SetValuePosition : Real;   // 正向运动的最大位置
            LU_Scale : Real;   // 默认--工程单位放大倍数
            p1520MaxFwdTorque : Real;   // 默认，最大正向扭矩，*基准扭矩
            p1521MaxBwdTorque : Real;   // 默认，最大负向向扭矩，*基准扭矩
            p2177MotorBlockedDelayTime : Real;   // 默认. 0.5秒
            p2634 : Real;   // 默认--扭矩模式时的跟随误差
            p2635 : Real;   // 默认--扭矩模式的监控范围，
            p2542_StaticMonitorError : Real;   // *_导程，即：默认静态监控误差为0.2*导程
            p2544_InpRange : Real;   // *_导程，即：默认静态监控误差为0.2*导程
            p2546FollowingError : Real;   // 默认--跟随误差
            p2572_P2573_AccDccTime : Real;   // 默认0.1S，按照0.1S时间加速到4800rpm计算加减速系数
            TimeOutSetValue : Time;   // 默认--15S内，命令必须能正常结束；
            ModularSettingValue : Real;   // 模态设定值
            sp : Array[0..3] of Real;   // 输入输出参数
            ConfigReference : Struct   // 输入输出参数
               SpeedOfSearchX8Ref_p2605 : Real;   // *_Unit: LU/S，找原点开关信号的速度，Exe 30.0mm/s
               SpeedOfSearchZeroMark_p2608 : Real;   // *_Unit: LU/S 找ZeroMark位置的速度Eg. 5.0mm/s
               SpeedOfMoveToZeroPos_p2611 : Real;   // *_Unit: LU/S，远点找到后的偏移速度Exe 60.0mm/s
               SpeedFast_Search_NoZeroMark : Real;   // *_Unit: *Lead/s. 不需要ZeroMark时的寻0速度
               SpeedSlow_Search_NoZeroMark : Real;   // *_Unit: *Lead/s. 不需要ZeroMark时的寻0速度
            END_STRUCT;
         END_STRUCT;
         Ref_Option : Struct   // 输入输出参数
            RefDirectionFwd : Bool;   // 1: 正向回原点，0：负向回原点；
            RefSource : Struct   // 原点开关的来源，只能有一个变量=On，否则后果自负
               op_CurrentPos : Bool;   // 当前位置作为原点
               op_X8_Ref_NO : Bool;   // 使用X8.DI1作为原点信号
               op_X8_Ref_NC : Bool;   // 使用取反后X8.DI1作为原点信号
               op_X8_CCWL : Bool;   // 使用X8.DI2负极限作为原点信号
               op_X8_CWL : Bool;   // 使用X8.DI3正极限作为原点信号
            END_STRUCT;
         END_STRUCT;
      END_STRUCT;
      Servo_CTRL_OUT : Struct   // 输入输出参数
         ActualPosition : Real;   // Actual Position (Directmode/Positioncontrol)
         ActualVelocity : Real;   // Actual Velocity %
         ParameterValue_DataCom : Real;   // Value of the parameter. Read Out from the controller
         MotorRatedTorque : Real;   // PNU1036.1,The motor's rated torque in 0.001 Nm.
         LastCylceTime : DInt;   // 动作时间
         Max_SetValueVelocity : Real;   // 计算得出的最大运动速度
         RecordComError : Int;   // Record Communication Error
         sp : Array[0..3] of Real;   // 输入输出参数
      END_STRUCT;
      Servo_Status : Struct   // 输入输出参数
         Busy : Bool;   // 运动控制循环调用中
         DataComBusy : Bool;   // 参数编辑循环调用中
         HomePos : Bool;   // 输出，已经回过原点
         WorkHomePos : Bool;   // 在工作原点
         TaskDone : Bool;   // 完成脉冲
         TaskIO : Bool;   // 命令执行异常结束
         TaskNIO : Bool;   // 命令执行异常结束
         DataComTaskDone : Bool;   // 通讯命令完成
         DataComTaskIO : Bool;   // 正常完成
         DataComTaskNIO : Bool;   // 异常完成
         OkToStart : Bool;   // 允许启动
         NotReady : Bool;   // 驱动器未就绪！
         FwdPmt : Bool;   // 前进允许_For TP Display
         BwdPmt : Bool;   // 后退允许_For TP Display
         TrackModePosDone : Bool;   // 定位命令下，位置已经到达
         ParameterInitOK : Bool;   // 输入输出参数
         TorqueLimited : Bool;   // 输入输出参数
         PromptValue : Int;   // 伺服状态
      END_STRUCT;
      sp : Array[1..24] of Byte;   // 备用
      IN : Bool;   // 输入输出参数
      Q : Bool;   // 输入输出参数
   END_VAR
   VAR
      TP_Cmd : Word := 30;   // 用于触摸屏传入命令
      TP_Status : Word;   // 用于Bit位的触摸屏显示
      Cmd : Struct   // 流程启动命令36
         Man : Struct   // 触摸屏内使用
            StartTest : Bool;   // 单循环测试
         END_STRUCT;
         Auto : Struct   // 触摸屏内使用
            StartTest : Bool;   // 单循环测试
         END_STRUCT;
         sp : Array[1..30] of Byte;   // 备用
      END_STRUCT;
      AtCmd : Struct   // 静态变量
         Man : Word;   // 静态变量
         Auto : Word;   // 静态变量
      END_STRUCT;
      Ctrl_IN : Struct   // 传入的参数_Start70
         TestCycleCounter : DInt := 1000000;   // 静态变量
         MinPos : Real := 10.0;   // 静态变量
         MaxPos : Real := 20.0;   // 静态变量
         InitParameter : Struct   // 静态变量
            TimeOutSetValue : Time := T#30S;   // 静态变量
            ServoTorque : Real := 0.4;   // 静态变量
            ServoVelocity : Real := 50.0;   // 静态变量
         END_STRUCT;
         sp : Array[1..16] of Byte;   // 备用
      END_STRUCT;
      Ctrl_Out : Struct   // 传出的数值结果_Start110
         AcutalCycleCounter : DInt;   // 静态变量
         LastCylceTime : DInt;   // 动作时间
         LastStep : Int;   // 静态变量
         sp : Array[1..30] of Byte;   // 备用
      END_STRUCT;
      Status : Struct   // 状态_Start150
         Busy : Bool;   // 主流程运行中
         OkToStart : Bool;   // 条件满足，允许启动
         sp : Bool;   // 静态变量
         sp_1 : Bool;   // 静态变量
         TaskDone : Bool;   // 静态变量
         TaskIO : Bool;   // 产品装配/测试后合格标志
         TaskNIO : Bool;   // 产品装配/测试后不合格标志
         PromptValue : Int;   // 伺服状态
      END_STRUCT;
      AtStatus : Word;   // 静态变量
      "Step" : Struct   // 过程步
         RandomStepNO : Word;   // 静态变量
         Main : Struct   // 运动控制步
            Start : Bool;   // 静态变量
            TimeOut : Bool;   // 静态变量
            ErrEnd : Bool;   // 静态变量
            End : Bool;   // 静态变量
            RandomTestCycleReStart : Bool;   // 静态变量
            S1 : Bool;   // 静态变量
            S2 : Bool;   // 静态变量
            S3 : Bool;   // 静态变量
            S4 : Bool;   // 静态变量
            S5 : Bool;   // 静态变量
            S6 : Bool;   // 静态变量
            S7 : Bool;   // 静态变量
            S8 : Bool;   // 静态变量
            S9 : Bool;   // 静态变量
            S10 : Bool;   // 静态变量
            S11 : Bool;   // 静态变量
            S12 : Bool;   // 静态变量
            S13 : Bool;   // 静态变量
            S14 : Bool;   // 静态变量
            S15 : Bool;   // 静态变量
            S16 : Bool;   // 静态变量
            S17 : Bool;   // 静态变量
            S18 : Bool;   // 静态变量
            S19 : Bool;   // 静态变量
            S20 : Bool;   // 静态变量
            S21 : Bool;   // 静态变量
            S22 : Bool;   // 静态变量
            S23 : Bool;   // 静态变量
            S24 : Bool;   // 静态变量
            S25 : Bool;   // 静态变量
            S26 : Bool;   // 静态变量
            S27 : Bool;   // 静态变量
            S28 : Bool;   // 静态变量
            S29 : Bool;   // 静态变量
            S30 : Bool;   // 静态变量
            S31 : Bool;   // 静态变量
            S32 : Bool;   // 静态变量
            S33 : Bool;   // 静态变量
            S34 : Bool;   // 静态变量
            S35 : Bool;   // 静态变量
            S36 : Bool;   // 静态变量
            S37 : Bool;   // 静态变量
            S38 : Bool;   // 静态变量
            S39 : Bool;   // 静态变量
            S40 : Bool;   // 静态变量
            S41 : Bool;   // 静态变量
            S42 : Bool;   // 静态变量
            S43 : Bool;   // 静态变量
            S44 : Bool;   // 静态变量
            S45 : Bool;   // 静态变量
            S46 : Bool;   // 静态变量
            S47 : Bool;   // 静态变量
            S48 : Bool;   // 静态变量
            S49 : Bool;   // 静态变量
            S50 : Bool;   // 静态变量
            S51 : Bool;   // 静态变量
            S52 : Bool;   // 静态变量
            S53 : Bool;   // 静态变量
            S54 : Bool;   // 静态变量
            S55 : Bool;   // 静态变量
            S56 : Bool;   // 静态变量
            S57 : Bool;   // 静态变量
            S58 : Bool;   // 静态变量
            S59 : Bool;   // 静态变量
            S60 : Bool;   // 静态变量
            S61 : Bool;   // 静态变量
            S62 : Bool;   // 静态变量
            DTResetS1 : Bool;   // 静态变量
            DTResetS2 : Bool;   // 静态变量
            DTResetS3 : Bool;   // 静态变量
            DTResetS4 : Bool;   // 静态变量
            DTResetS5 : Bool;   // 静态变量
            DTResetS6 : Bool;   // 静态变量
            DTResetS7 : Bool;   // 静态变量
            DTResetS8 : Bool;   // 静态变量
         END_STRUCT;
      END_STRUCT;
      InfoStruct : Struct   // 信息
         Stopped : Bool;   // A00. Controller Stopped
         Halt : Bool;   // A01. Controller Halt
         WaitForTargetPosReached : Bool;   // A02. Wait for targetPos Reached!
         WaitForTargetPosInBand : Bool;   // A03. Wait for target pos in Band!
         ModeOff : Bool;   // A04. ModeOff !
         StartProhibit : Bool;   // A05. Permit = off
         Ready : Bool;   // A06. Ready to start
         AlarmPresent : Bool;   // A07. Alarm Present
         WaitForStandStill : Bool;   // A10. Wait for StandStil (check p1226 )
         FwdNotPmt : Bool;   // A11. forbid axis to forward !
         BwdNotPmt : Bool;   // A12. forbid axis to backward !
         StartHoming : Bool;   // A13. Home Seek Started
         StartWorkHome : Bool;   // A14. Start Work home process
         StartTaskPos : Bool;   // A15. Start Position process!
         StartTraversingBlock : Bool;   // A16. StartTraversingBlock
         StartJog : Bool;   // A17. Start Jog movement
         StartTorqueCtrlMode : Bool;   // A20. Start Torque Control Mode
         DataComExecuting : Bool;   // A21. Executing parameter communication..
         TrackingModeActive : Bool;   // A22. TrackIngModeActive
         LeavingReference : Bool;   // A23. Ref = ON, Leaving away Ref Pos !
         sp31 : Bool;   // A24.
         sp33 : Bool;   // A25.
         sp34 : Bool;   // A26.
         sp35 : Bool;   // A27.
         sp36 : Bool;   // A30.
         x : Bool;   // A31
         x_1 : Bool;   // A32
         x_2 : Bool;   // A33
         x_3 : Bool;   // A34
         x_4 : Bool;   // A35
         x_5 : Bool;   // A36
         x_6 : Bool;   // A37
      END_STRUCT;
      ErrStruct : Struct   // 故障
         DPConnectErr : Bool;   // E00. Connnect Err, Pls Reset!
         DriveDisableByUser : Bool;   // E01. DriveDisabled by user
         InitPara : Bool;   // E02. PLC is sending init para to Drive!
         ControlViaPLCError : Bool;   // E03. Control via PLC Error, Pls check V-Assistant
         DriveNotReadyForSwitchON : Bool;   // E04. Drive Not Ready For Switch ON, Check DC Supply
         DriveEnableFail : Bool;   // E05. Drive Enable Failue
         FaultPresent : Bool;   // E06. Fault Present !
         ReferenceFail : Bool;   // E07. Reference sensor fault, pls check !
         RecordComError : Bool;   // E10. Record Communication Error
         EndofMotionError : Bool;   // E11. End of Motion fault present
         EndOfTimeOut : Bool;   // E12. Cmd end of time Out !
         CWL_Approached : Bool;   // E13. Controller X8.DI3.CWL = Off, pls Check !
         CCWL_Approached : Bool;   // E14. Controller X8.DI2.CCWL = Off, pls Check!
         RefSourceNotSet : Bool;   // E15.CTRL_IN.RefSource not set !
         EMOKError : Bool;   // E16. X8.DI4.EMOK = Off,pls Check !
         SetValuePos_MinError : Bool;   // E17. SetValuePosition too small !
         AdjustFail_Counter : Bool;   // E20. Adjust fail, counter is finished
         AdjustFail_FlowRateLow : Bool;   // E21. Adjust fail, FlowRate is too low !
         sp31 : Bool;   // E22
         sp33 : Bool;   // E23
         sp34 : Bool;   // E24
         sp35 : Bool;   // E25
         sp36 : Bool;   // E26
         sp37 : Bool;   // E27
         xx_8 : Bool;   // E30
         xx_9 : Bool;   // E31
         xx_10 : Bool;   // E32
         xx_11 : Bool;   // E33
         xx_12 : Bool;   // E34
         sp32 : Bool;   // E35
         sp38 : Bool;   // E36
         sp39 : Bool;   // E37
      END_STRUCT;
      FB_InfoPrompt : "FB1021_Prompt_Object";   // 信息
      FB_ErrPrompt : "FB1021_Prompt_Object";   // 故障
      Timer_TimeOut : "FB950_SDTimer";   // 静态变量
      Aux : Struct   // 静态变量
         CycleTime_StartTime : DInt;   // 开始循环的时间
         TimeOutSetValue : Time;   // 默认--15S内，命令必须能正常结束；
         sp : Array[1..278] of Byte;   // 静态变量
      END_STRUCT;
      LastAddr : Int := 498;   // 总占地址
      CycleTime : Int;   // 静态变量
      PromptValueBake : Int;   // 静态变量
      ShiftBake : Int;   // 静态变量
      TempSystime : Time;   // 静态变量
   END_VAR
   VAR_TEMP
      AnyCmdOn : Bool;   // 临时变量
      T_int : Int;   // 临时变量
      T_RetVal : Int;   // 临时变量
      T_DINT : DInt;   // 临时变量
      T_Real : Real;   // 临时变量
      VolTargetMin : Real;   // 临时变量
      VolTargetMax : Real;   // 临时变量
      Tol_Min_PartDP : Real;   // 临时变量
      Tol_Max_PartDP : Real;   // 临时变量
   END_VAR
BEGIN

   // ---------- 网络 1 ----------
   // 标题：<<<触摸屏使用的变量传递
   // 含义：将 #TP_Cmd 赋给 #AtCmd.Man
   #AtCmd.Man := #TP_Cmd;
   // 含义：将 #AtStatus 赋给 #TP_Status
   #TP_Status := #AtStatus;
   // 含义：条件 NOT (#AllMode) 成立时，将 0 传送到 #TP_Cmd
   IF NOT (#AllMode) THEN
       #TP_Cmd := 0;
   END_IF;

   // ---------- 网络 2 ----------
   // 标题：E12. Cmd end of time Out !
   // 含义：条件 #ErrRst 成立时，将 FALSE 传送到 #ErrStruct.EndOfTimeOut
   IF #ErrRst THEN
       #ErrStruct.EndOfTimeOut := FALSE;
   END_IF;

